(* IEC 61131-3 sources: daoli-st-library/DL_Base (part 6) *)

(* ---- FC_DL_MapRangeIntQuant.st ---- *)
(*
  FC_DL_MapRangeIntQuant —— 量程映射加整数量化，步长加四舍五入
  分类：DL_Base | 复杂度：2 | 轮次：R86
  开源溯源：道莅原创（clean-room 自研，纯 IEC 61131-3 通用算法），无外部代码引用
  许可证：MIT
  职责：先把输入线性映射到输出量程（输入越界钳位），再按 fStep 步长量化到整数刻度：
        nTick = round(mapped / step)，fOut = nTick * step；fTick 为量化后的整数刻度。
  契约：fIn 输入、fInMin/fInMax 输入端点、fOutMin/fOutMax 输出端点、fStep 步长（必须 > 0）；
        fOut 量化结果 [输出量程单位]、fTick 整数刻度；返回 TRUE 表示可信。
  边界：① 步长零 / 负值前置判（除零防护）；② 量程退化校验（容差 DL_MQ_EPS）；
        ③ 六个浮点入参逐一非有限闸；④ 转整前对刻度做 ±1.0E6 上限兜底，避免 LREAL_TO_DINT 越域；
        ⑤ 零全局、零物理地址、零库件依赖。
*)
FUNCTION FC_DL_MapRangeIntQuant : BOOL
VAR_INPUT
    fIn     : LREAL := 0.0;            // 输入值 [输入量程单位] / The input value
    fInMin  : LREAL := 0.0;            // 输入量程下端点 [输入量程单位] / The input range low end
    fInMax  : LREAL := 100.0;          // 输入量程上端点 [输入量程单位] / The input range high end
    fOutMin : LREAL := 0.0;            // 输出量程下端点 [输出量程单位] / The output range low end
    fOutMax : LREAL := 100.0;          // 输出量程上端点 [输出量程单位] / The output range high end
    fStep   : LREAL := 1.0;            // 量化步长（必须 > 0） [输出量程单位] / The quantisation step
END_VAR
VAR_OUTPUT
    fOut  : LREAL;                     // 量化后的结果 [输出量程单位] / The quantised result
    fTick : LREAL;                     // 量化后的整数刻度值 [刻度] / The integer tick value as a real
END_VAR
VAR
    xBad     : BOOL;                   // 参数非法标志 [—] / The parameter invalid flag
    fInSpan  : LREAL;                  // 输入量程跨度 [输入量程单位] / The input span
    fMapped  : LREAL;                  // 未量化的映射值 [输出量程单位] / The mapped value
    fTicks   : LREAL;                  // 未取整的刻度 [刻度] / The raw tick count
    diTick   : DINT;                   // 四舍五入后的整数刻度 [刻度] / The rounded tick count
END_VAR
VAR CONSTANT
    DL_MQ_EPS  : LREAL := 1.0E-9;      // 浮点比较容差 [-] / The floating point comparison tolerance
    DL_MQ_INF  : LREAL := 1.0E30;      // 非有限 / 越界判据上限 [-] / The magnitude gate
    DL_MQ_TICK : LREAL := 1.0E6;       // 转整前的刻度上限兜底 [刻度] / The tick guard before conversion
    DL_MQ_HALF : LREAL := 0.5;         // 四舍五入偏置 [-] / The rounding bias
    DL_MQ_Z    : LREAL := 0.0;         // 浮点零常量 [-] / The floating point zero constant
END_VAR

FC_DL_MapRangeIntQuant := FALSE;                          // 返回值预置假 / preset the return false
fOut := fOutMin;                                          // 输出预置为输出下端点哨兵 / preset the low end sentinel
fTick := DL_MQ_Z;                                         // 刻度预置零 [刻度] / preset the tick zero
xBad := FALSE;                                            // 非法标志预置假 / preset the invalid flag false
IF (fIn <> fIn) OR (ABS(fIn) > DL_MQ_INF) THEN            // 输入非有限闸 / the input gate
    xBad := TRUE;                                         // 置非法标志 / raise the invalid flag
END_IF
IF (fInMin <> fInMin) OR (ABS(fInMin) > DL_MQ_INF) THEN   // 输入下端非有限闸 / the input low end gate
    xBad := TRUE;                                         // 置非法标志 / raise the invalid flag
END_IF
IF (fInMax <> fInMax) OR (ABS(fInMax) > DL_MQ_INF) THEN   // 输入上端非有限闸 / the input high end gate
    xBad := TRUE;                                         // 置非法标志 / raise the invalid flag
END_IF
IF (fOutMin <> fOutMin) OR (ABS(fOutMin) > DL_MQ_INF) THEN // 输出下端非有限闸 / the output low end gate
    xBad := TRUE;                                         // 置非法标志 / raise the invalid flag
END_IF
IF (fOutMax <> fOutMax) OR (ABS(fOutMax) > DL_MQ_INF) THEN // 输出上端非有限闸 / the output high end gate
    xBad := TRUE;                                         // 置非法标志 / raise the invalid flag
END_IF
IF (fStep <> fStep) OR (ABS(fStep) > DL_MQ_INF) THEN      // 步长非有限闸 / the step gate
    xBad := TRUE;                                         // 置非法标志 / raise the invalid flag
END_IF
IF fStep <= DL_MQ_EPS THEN                                // 步长非正（除零防护） / the step is not positive
    xBad := TRUE;                                         // 置非法标志 / raise the invalid flag
END_IF
fInSpan := fInMax - fInMin;                               // 输入量程跨度 [输入量程单位] / the input span
IF ABS(fInSpan) < DL_MQ_EPS THEN                          // 输入量程退化（除零防护） / the degenerate input span
    xBad := TRUE;                                         // 置非法标志 / raise the invalid flag
END_IF
IF NOT xBad THEN                                          // 参数全通过才映射量化 / map and quantise when all pass
    fMapped := fIn;                                       // 输入接管 [输入量程单位] / take the input value
    IF fInSpan > DL_MQ_Z THEN                             // 正常量程方向 / the normal direction
        IF fMapped < fInMin THEN                          // 低于下端点 / below the low end
            fMapped := fInMin;                            // 钳到下端点 [输入量程单位] / clamp to the low end
        END_IF
        IF fMapped > fInMax THEN                          // 高于上端点 / above the high end
            fMapped := fInMax;                            // 钳到上端点 [输入量程单位] / clamp to the high end
        END_IF
    ELSE                                                  // 反向量程 / the reversed direction
        IF fMapped > fInMin THEN                          // 高于下端点 / above the low end
            fMapped := fInMin;                            // 钳到下端点 [输入量程单位] / clamp to the low end
        END_IF
        IF fMapped < fInMax THEN                          // 低于上端点 / below the high end
            fMapped := fInMax;                            // 钳到上端点 [输入量程单位] / clamp to the high end
        END_IF
    END_IF
    fMapped := fOutMin + ((fMapped - fInMin) / fInSpan) * (fOutMax - fOutMin); // 线性映射（分母已证非零）
    fTicks := fMapped / fStep;                            // 换算成刻度数（步长已证正） [刻度] / the raw tick count
    IF fTicks > DL_MQ_TICK THEN                           // 刻度上越界，转整前兜底 / the positive tick guard
        fTicks := DL_MQ_TICK;                             // 钳到刻度上限 [刻度] / clamp the tick count
    END_IF
    IF fTicks < -DL_MQ_TICK THEN                          // 刻度下越界，转整前兜底 / the negative tick guard
        fTicks := -DL_MQ_TICK;                            // 钳到刻度下限 [刻度] / clamp the tick count
    END_IF
    IF fTicks >= DL_MQ_HALF THEN                          // 非负四舍五入 / non negative rounding
        diTick := LREAL_TO_DINT(fTicks + DL_MQ_HALF);     // 加半后截断 [刻度] / add a half then truncate
    ELSIF fTicks <= -DL_MQ_HALF THEN                      // 非正四舍五入 / non positive rounding
        diTick := LREAL_TO_DINT(fTicks - DL_MQ_HALF);     // 减半后截断 [刻度] / subtract a half then truncate
    ELSE
        diTick := 0;                                      // 近零带归零 [刻度] / the near zero band
    END_IF
    fTick := DINT_TO_LREAL(diTick);                       // 整数刻度出口 [刻度] / publish the integer tick
    fOut := fTick * fStep;                                // 量化结果还原 [输出量程单位] / restore the quantised value
    FC_DL_MapRangeIntQuant := TRUE;                       // 量化成功 / the quantisation succeeded
ELSE
    fOut := fOutMin;                                      // 非法参数输出下端点哨兵 [输出量程单位] / the sentinel
    fTick := DL_MQ_Z;                                     // 刻度输出零哨兵 [刻度] / the tick sentinel
    FC_DL_MapRangeIntQuant := FALSE;                      // 结果不可信 / the result is not valid
END_IF
END_FUNCTION

(* ---- FC_DL_MapRangeInverseSolve.st ---- *)
(*
  FC_DL_MapRangeInverseSolve —— 由工程值反解原始量程值，含钳位
  分类：DL_Base | 复杂度：2 | 轮次：R86
  开源溯源：道莅原创（clean-room 自研，纯 IEC 61131-3 通用算法），无外部代码引用
  许可证：MIT
  职责：正向映射 out = fOutMin + (in - fInMin)/(fInMax - fInMin) * (fOutMax - fOutMin) 的逆解：
        raw = fInMin + (fOut - fOutMin) * (fInMax - fInMin) / (fOutMax - fOutMin)。
  契约：fEng 工程值输入 [输出量程单位]、fInMin/fInMax 原始量程端点、fOutMin/fOutMax 工程量程端点；
        fRaw 反解结果 [原始量程单位]（钳在原始量程内）；返回 TRUE 表示可信。
  边界：① 除零防护：分母 fOutSpan 过退化闸后才做除法；② 反解结果按原始量程钳位；
        ③ 五个浮点入参逐一非有限闸；④ 零全局、零物理地址、零库件依赖。
*)
FUNCTION FC_DL_MapRangeInverseSolve : BOOL
VAR_INPUT
    fEng    : LREAL := 0.0;            // 工程值输入 [输出量程单位] / The engineering value input
    fInMin  : LREAL := 0.0;            // 原始量程下端点 [原始量程单位] / The raw range low end
    fInMax  : LREAL := 100.0;          // 原始量程上端点 [原始量程单位] / The raw range high end
    fOutMin : LREAL := 0.0;            // 工程量程下端点 [输出量程单位] / The engineering range low end
    fOutMax : LREAL := 100.0;          // 工程量程上端点 [输出量程单位] / The engineering range high end
END_VAR
VAR_OUTPUT
    fRaw : LREAL;                      // 反解结果 [原始量程单位] / The solved raw value
END_VAR
VAR
    xBad      : BOOL;                  // 参数非法标志 [—] / The parameter invalid flag
    fEngClamp : LREAL;                 // 钳位后的工程值 [输出量程单位] / The clamped engineering value
    fOutSpan  : LREAL;                 // 工程量程跨度 [输出量程单位] / The engineering span
    fInSpan   : LREAL;                 // 原始量程跨度 [原始量程单位] / The raw span
    fRawCalc  : LREAL;                 // 未钳位的反解结果 [原始量程单位] / The unclamped solved value
END_VAR
VAR CONSTANT
    DL_MI_EPS : LREAL := 1.0E-9;       // 浮点比较容差 [-] / The floating point comparison tolerance
    DL_MI_INF : LREAL := 1.0E30;       // 非有限 / 越界判据上限 [-] / The magnitude gate
    DL_MI_Z   : LREAL := 0.0;          // 浮点零常量 [-] / The floating point zero constant
END_VAR

FC_DL_MapRangeInverseSolve := FALSE;                      // 返回值预置假 / preset the return false
fRaw := fInMin;                                           // 输出预置为原始量程下端点哨兵 / preset the raw low end sentinel
xBad := FALSE;                                            // 非法标志预置假 / preset the invalid flag false
IF (fEng <> fEng) OR (ABS(fEng) > DL_MI_INF) THEN         // 工程值非有限闸 / the engineering value gate
    xBad := TRUE;                                         // 置非法标志 / raise the invalid flag
END_IF
IF (fInMin <> fInMin) OR (ABS(fInMin) > DL_MI_INF) THEN   // 原始下端非有限闸 / the raw low end gate
    xBad := TRUE;                                         // 置非法标志 / raise the invalid flag
END_IF
IF (fInMax <> fInMax) OR (ABS(fInMax) > DL_MI_INF) THEN   // 原始上端非有限闸 / the raw high end gate
    xBad := TRUE;                                         // 置非法标志 / raise the invalid flag
END_IF
IF (fOutMin <> fOutMin) OR (ABS(fOutMin) > DL_MI_INF) THEN // 工程下端非有限闸 / the engineering low end gate
    xBad := TRUE;                                         // 置非法标志 / raise the invalid flag
END_IF
IF (fOutMax <> fOutMax) OR (ABS(fOutMax) > DL_MI_INF) THEN // 工程上端非有限闸 / the engineering high end gate
    xBad := TRUE;                                         // 置非法标志 / raise the invalid flag
END_IF
fOutSpan := fOutMax - fOutMin;                            // 工程量程跨度 [输出量程单位] / the engineering span
fInSpan := fInMax - fInMin;                               // 原始量程跨度 [原始量程单位] / the raw span
IF ABS(fOutSpan) < DL_MI_EPS THEN                         // 工程跨度退化（除零防护） / the degenerate engineering span
    xBad := TRUE;                                         // 置非法标志 / raise the invalid flag
END_IF
IF NOT xBad THEN                                          // 参数全通过才反解 / solve only when all parameters pass
    fEngClamp := fEng;                                    // 工程值接管 [输出量程单位] / take the engineering value
    IF fOutSpan > DL_MI_Z THEN                            // 正常方向 / the normal direction
        IF fEngClamp < fOutMin THEN                       // 低于工程下端点 / below the engineering low end
            fEngClamp := fOutMin;                         // 钳到工程下端点 [输出量程单位] / clamp to the low end
        END_IF
        IF fEngClamp > fOutMax THEN                       // 高于工程上端点 / above the engineering high end
            fEngClamp := fOutMax;                         // 钳到工程上端点 [输出量程单位] / clamp to the high end
        END_IF
    ELSE                                                  // 反向工程跨度 / the reversed engineering span
        IF fEngClamp > fOutMin THEN                       // 高于工程下端点 / above the engineering low end
            fEngClamp := fOutMin;                         // 钳到工程下端点 [输出量程单位] / clamp to the low end
        END_IF
        IF fEngClamp < fOutMax THEN                       // 低于工程上端点 / below the engineering high end
            fEngClamp := fOutMax;                         // 钳到工程上端点 [输出量程单位] / clamp to the high end
        END_IF
    END_IF
    fRawCalc := fInMin + ((fEngClamp - fOutMin) / fOutSpan) * fInSpan; // 反解（分母已证非零） [原始量程单位]
    IF fInMax >= fInMin THEN                              // 原始量程正常方向 / the normal raw direction
        IF fRawCalc < fInMin THEN                         // 反解低于原始下端点 / below the raw low end
            fRawCalc := fInMin;                           // 钳到原始下端点 [原始量程单位] / clamp to the low end
        END_IF
        IF fRawCalc > fInMax THEN                         // 反解高于原始上端点 / above the raw high end
            fRawCalc := fInMax;                           // 钳到原始上端点 [原始量程单位] / clamp to the high end
        END_IF
    ELSE                                                  // 原始量程反向 / the reversed raw range
        IF fRawCalc > fInMin THEN                         // 反解高于原始下端点 / above the raw low end
            fRawCalc := fInMin;                           // 钳到原始下端点 [原始量程单位] / clamp to the low end
        END_IF
        IF fRawCalc < fInMax THEN                         // 反解低于原始上端点 / below the raw high end
            fRawCalc := fInMax;                           // 钳到原始上端点 [原始量程单位] / clamp to the high end
        END_IF
    END_IF
    fRaw := fRawCalc;                                     // 反解结果出口 [原始量程单位] / publish the solved value
    FC_DL_MapRangeInverseSolve := TRUE;                   // 反解成功 / the solve succeeded
ELSE
    fRaw := fInMin;                                       // 非法参数输出原始下端点哨兵 [原始量程单位] / the sentinel
    FC_DL_MapRangeInverseSolve := FALSE;                  // 结果不可信 / the result is not valid
END_IF
END_FUNCTION

(* ---- FC_DL_MapRangePiecewise3.st ---- *)
(*
  FC_DL_MapRangePiecewise3 —— 三段折线映射，分段斜率加断点连续校验
  分类：DL_Base | 复杂度：2 | 轮次：R86
  开源溯源：道莅原创（clean-room 自研，纯 IEC 61131-3 通用算法），无外部代码引用
  许可证：MIT
  职责：由 4 个断点（afX 单调递增）与对应 4 个输出值构造三段折线，按输入落在哪一段做线性插值；
        断点单调性即保证折线在断点处连续（左段右端值 = 右段左端值 = afY[i]）。
  契约：fIn 输入、afX 断点横坐标（必须严格递增）、afY 断点纵坐标；fOut 折线输出；返回 TRUE 表示可信。
  边界：① 断点严格递增校验（容差 DL_MW_EPS），否则判非法；② 所有断点与输入做非有限闸；
        ③ 输入越两端断点时钳到端点（不外插）；④ 除零防护：段跨度经单调性闸后恒 > 0；
        ⑤ 零全局、零物理地址、零库件依赖；数组为显式定长（R15）。
*)
FUNCTION FC_DL_MapRangePiecewise3 : BOOL
VAR_INPUT
    fIn  : LREAL := 0.0;                             // 输入值 [输入量程单位] / The input value
    afX  : ARRAY[0..3] OF LREAL;                     // 四个断点横坐标（严格递增） [输入量程单位] / The breakpoints
    afY  : ARRAY[0..3] OF LREAL;                     // 四个断点纵坐标 [输出量程单位] / The breakpoint outputs
END_VAR
VAR_OUTPUT
    fOut  : LREAL;                                   // 折线输出 [输出量程单位] / The piecewise output
    nSeg  : INT;                                     // 命中段号（0..2） [下标] / The hit segment index
END_VAR
VAR
    xBad  : BOOL;                                    // 参数非法标志 [—] / The parameter invalid flag
    xFound : BOOL;                                   // 命中段查找标志 [—] / The hit segment search flag
    i     : INT;                                     // 遍历索引 [下标] / The traversal index
    k     : INT;                                     // 命中段索引 [下标] / The hit segment index
    fSpan : LREAL;                                   // 命中段的横坐标跨度 [输入量程单位] / The segment span
END_VAR
VAR CONSTANT
    DL_MW_EPS  : LREAL := 1.0E-9;                    // 浮点比较容差 [-] / The floating point comparison tolerance
    DL_MW_INF  : LREAL := 1.0E30;                    // 非有限 / 越界判据上限 [-] / The magnitude gate
    DL_MW_Z    : LREAL := 0.0;                       // 浮点零常量 [-] / The floating point zero constant
    DL_MW_N    : INT := 3;                           // 折线段数 [段] / The number of segments
    DL_MW_I0   : INT := 0;                           // 下标零 [下标] / The index zero
END_VAR

FC_DL_MapRangePiecewise3 := FALSE;                    // 返回值预置假 / preset the return false
fOut := DL_MW_Z;                                      // 输出预置零哨兵 / preset the zero sentinel
nSeg := DL_MW_I0;                                     // 段号预置零 [下标] / preset the segment index zero
xBad := FALSE;                                        // 非法标志预置假 / preset the invalid flag false
IF (fIn <> fIn) OR (ABS(fIn) > DL_MW_INF) THEN        // 输入非有限闸 / the input gate
    xBad := TRUE;                                     // 置非法标志 / raise the invalid flag
END_IF
FOR i := DL_MW_I0 TO DL_MW_N DO                       // 四个断点逐一校验 / check every breakpoint
    IF (afX[i] <> afX[i]) OR (ABS(afX[i]) > DL_MW_INF) THEN // 横坐标非有限 / the abscissa is not finite
        xBad := TRUE;                                 // 置非法标志 / raise the invalid flag
    END_IF
    IF (afY[i] <> afY[i]) OR (ABS(afY[i]) > DL_MW_INF) THEN // 纵坐标非有限 / the ordinate is not finite
        xBad := TRUE;                                 // 置非法标志 / raise the invalid flag
    END_IF
END_FOR
FOR i := DL_MW_I0 TO DL_MW_N - 1 DO                   // 相邻断点严格递增校验 / strictly increasing check
    IF (afX[i + 1] - afX[i]) < DL_MW_EPS THEN         // 跨度非正（含重合断点） / a non positive span
        xBad := TRUE;                                 // 置非法标志 / raise the invalid flag
    END_IF
END_FOR
IF NOT xBad THEN                                      // 参数全通过才插值 / interpolate when all parameters pass
    IF fIn <= afX[DL_MW_I0] THEN                      // 低于最低断点，钳到端点 / below the lowest breakpoint
        fOut := afY[DL_MW_I0];                        // 取最低断点输出 [输出量程单位] / take the lowest output
        nSeg := DL_MW_I0;                             // 段号记零 [下标] / the segment index is zero
    ELSIF fIn >= afX[DL_MW_N] THEN                    // 高于最高断点，钳到端点 / above the highest breakpoint
        fOut := afY[DL_MW_N];                         // 取最高断点输出 [输出量程单位] / take the highest output
        nSeg := DL_MW_N - 1;                          // 段号记末段 [下标] / the last segment index
    ELSE
        k := DL_MW_I0;                                // 段索引从零起 / the segment index starts at zero
        xFound := FALSE;                              // 命中标志预置假 / preset the hit flag false
        WHILE (k <= DL_MW_N - 1) AND NOT xFound DO    // 显式递增查找命中段（有界） / find the hit segment
            IF fIn < afX[k + 1] THEN                  // 落在第 k 段内 / inside the k th segment
                xFound := TRUE;                       // 置命中标志 / raise the hit flag
            ELSE
                k := k + 1;                           // 继续下一段 / advance to the next segment
            END_IF
        END_WHILE
        IF k > DL_MW_N - 1 THEN                       // 命中段上越界兜底 / the hit index fallback
            k := DL_MW_N - 1;                         // 钳到末段 [下标] / clamp to the last segment
        END_IF
        fSpan := afX[k + 1] - afX[k];                 // 命中段跨度（已证 > 容差） [输入量程单位] / the segment span
        fOut := afY[k] + ((fIn - afX[k]) / fSpan) * (afY[k + 1] - afY[k]); // 段内线性插值 [输出量程单位]
        nSeg := k;                                    // 段号出口 [下标] / publish the hit segment
    END_IF
    FC_DL_MapRangePiecewise3 := TRUE;                 // 插值成功 / the interpolation succeeded
ELSE
    fOut := DL_MW_Z;                                  // 非法参数输出零哨兵 [输出量程单位] / the sentinel
    FC_DL_MapRangePiecewise3 := FALSE;                // 结果不可信 / the result is not valid
END_IF
END_FUNCTION

(* ---- FC_DL_MapRangeSatOut.st ---- *)
(*
  FC_DL_MapRangeSatOut —— 输入量程映射后对输出独立饱和限幅
  分类：DL_Base | 复杂度：2 | 轮次：R86
  开源溯源：道莅原创（clean-room 自研，纯 IEC 61131-3 通用算法），无外部代码引用
  许可证：MIT
  职责：先做 [fInMin, fInMax] → [fOutMin, fOutMax] 的线性映射（输入先钳到量程），
        再把映射结果独立钳到执行机构允许的 [fSatMin, fSatMax]（该区间可比输出量程更窄）。
  契约：fIn 输入、fInMin/fInMax 输入端点、fOutMin/fOutMax 输出端点、fSatMin/fSatMax 输出饱和限；
        fOut 结果；xSat 报告输出侧发生饱和；返回 TRUE 表示可信。
  边界：① 输入量程与饱和区间双退化校验（容差 DL_MS_EPS）；② 八个浮点入参逐一非有限闸；
        ③ 除零防护：除以 fInSpan 前已过退化闸；④ 零全局、零物理地址、零库件依赖。
*)
FUNCTION FC_DL_MapRangeSatOut : BOOL
VAR_INPUT
    fIn     : LREAL := 0.0;            // 输入值 [输入量程单位] / The input value
    fInMin  : LREAL := 0.0;            // 输入量程下端点 [输入量程单位] / The input range low end
    fInMax  : LREAL := 100.0;          // 输入量程上端点 [输入量程单位] / The input range high end
    fOutMin : LREAL := 0.0;            // 输出量程下端点 [输出量程单位] / The output range low end
    fOutMax : LREAL := 100.0;          // 输出量程上端点 [输出量程单位] / The output range high end
    fSatMin : LREAL := 0.0;            // 输出饱和下限 [输出量程单位] / The output saturation low limit
    fSatMax : LREAL := 100.0;          // 输出饱和上限 [输出量程单位] / The output saturation high limit
END_VAR
VAR_OUTPUT
    fOut : LREAL;                      // 结果（含输出侧饱和） [输出量程单位] / The saturated result
    xSat : BOOL;                       // 输出侧发生饱和 [—] / The output stage saturated
END_VAR
VAR
    xBad      : BOOL;                  // 参数非法标志 [—] / The parameter invalid flag
    fInClamp  : LREAL;                 // 钳位后的输入 [输入量程单位] / The clamped input
    fInSpan   : LREAL;                 // 输入量程跨度 [输入量程单位] / The input span
    fMapped   : LREAL;                 // 未限幅的映射结果 [输出量程单位] / The mapped value before limiting
END_VAR
VAR CONSTANT
    DL_MS_EPS : LREAL := 1.0E-9;       // 浮点比较容差 [-] / The floating point comparison tolerance
    DL_MS_INF : LREAL := 1.0E30;       // 非有限 / 越界判据上限 [-] / The magnitude gate
    DL_MS_Z   : LREAL := 0.0;          // 浮点零常量 [-] / The floating point zero constant
END_VAR

FC_DL_MapRangeSatOut := FALSE;                            // 返回值预置假 / preset the return false
fOut := fOutMin;                                          // 输出预置为输出下端点哨兵 / preset the low end sentinel
xSat := FALSE;                                            // 饱和标志预置假 / preset the saturation flag false
xBad := FALSE;                                            // 非法标志预置假 / preset the invalid flag false
IF (fIn <> fIn) OR (ABS(fIn) > DL_MS_INF) THEN            // 输入非有限闸 / the input gate
    xBad := TRUE;                                         // 置非法标志 / raise the invalid flag
END_IF
IF (fInMin <> fInMin) OR (ABS(fInMin) > DL_MS_INF) THEN   // 输入下端非有限闸 / the input low end gate
    xBad := TRUE;                                         // 置非法标志 / raise the invalid flag
END_IF
IF (fInMax <> fInMax) OR (ABS(fInMax) > DL_MS_INF) THEN   // 输入上端非有限闸 / the input high end gate
    xBad := TRUE;                                         // 置非法标志 / raise the invalid flag
END_IF
IF (fOutMin <> fOutMin) OR (ABS(fOutMin) > DL_MS_INF) THEN // 输出下端非有限闸 / the output low end gate
    xBad := TRUE;                                         // 置非法标志 / raise the invalid flag
END_IF
IF (fOutMax <> fOutMax) OR (ABS(fOutMax) > DL_MS_INF) THEN // 输出上端非有限闸 / the output high end gate
    xBad := TRUE;                                         // 置非法标志 / raise the invalid flag
END_IF
IF (fSatMin <> fSatMin) OR (ABS(fSatMin) > DL_MS_INF) THEN // 饱和下限非有限闸 / the saturation low gate
    xBad := TRUE;                                         // 置非法标志 / raise the invalid flag
END_IF
IF (fSatMax <> fSatMax) OR (ABS(fSatMax) > DL_MS_INF) THEN // 饱和上限非有限闸 / the saturation high gate
    xBad := TRUE;                                         // 置非法标志 / raise the invalid flag
END_IF
fInSpan := fInMax - fInMin;                               // 输入量程跨度 [输入量程单位] / the input span
IF ABS(fInSpan) < DL_MS_EPS THEN                          // 输入量程退化（除零防护） / the degenerate input span
    xBad := TRUE;                                         // 置非法标志 / raise the invalid flag
END_IF
IF fSatMax < fSatMin THEN                                 // 饱和区间倒置 / the saturated band is inverted
    xBad := TRUE;                                         // 置非法标志 / raise the invalid flag
END_IF
IF NOT xBad THEN                                          // 参数全通过才映射 / map only when all parameters pass
    fInClamp := fIn;                                      // 输入接管 [输入量程单位] / take the input value
    IF fInSpan > DL_MS_Z THEN                             // 正常量程方向 / the normal direction
        IF fInClamp < fInMin THEN                         // 低于下端点 / below the low end
            fInClamp := fInMin;                           // 钳到下端点 [输入量程单位] / clamp to the low end
        END_IF
        IF fInClamp > fInMax THEN                         // 高于上端点 / above the high end
            fInClamp := fInMax;                           // 钳到上端点 [输入量程单位] / clamp to the high end
        END_IF
    ELSE                                                  // 反向量程 / the reversed direction
        IF fInClamp > fInMin THEN                         // 高于下端点 / above the low end
            fInClamp := fInMin;                           // 钳到下端点 [输入量程单位] / clamp to the low end
        END_IF
        IF fInClamp < fInMax THEN                         // 低于上端点 / below the high end
            fInClamp := fInMax;                           // 钳到上端点 [输入量程单位] / clamp to the high end
        END_IF
    END_IF
    fMapped := fOutMin + ((fInClamp - fInMin) / fInSpan) * (fOutMax - fOutMin); // 线性映射（分母已证非零）
    fOut := fMapped;                                      // 映射值接入输出侧限幅 [输出量程单位] / take the mapped value
    IF fMapped > fSatMax THEN                             // 输出侧上饱和 / the output stage saturates high
        fOut := fSatMax;                                  // 钳到饱和上限 [输出量程单位] / clamp to the high limit
        xSat := TRUE;                                     // 置饱和标志 [—] / raise the saturation flag
    END_IF
    IF fMapped < fSatMin THEN                             // 输出侧下饱和 / the output stage saturates low
        fOut := fSatMin;                                  // 钳到饱和下限 [输出量程单位] / clamp to the low limit
        xSat := TRUE;                                     // 置饱和标志 [—] / raise the saturation flag
    END_IF
    FC_DL_MapRangeSatOut := TRUE;                         // 映射成功 / the mapping succeeded
ELSE
    fOut := fOutMin;                                      // 非法参数输出下端点哨兵 [输出量程单位] / the sentinel
    FC_DL_MapRangeSatOut := FALSE;                        // 结果不可信 / the result is not valid
END_IF
END_FUNCTION

(* ---- FC_DL_MaskCompare.st ---- *)
(*==============================================================================
 * 组件名称 (Component)  : FC_DL_MaskCompare
 * 所属子库 (Sublibrary) : DL_Base
 * 归属目录 (Directory)  : C:\Library\DL_Base
 * 当前版本 (Version)    : 1.0.0
 * 分类/来源标签         : 函数（FUNCTION）· 纯函数 · 状态字掩码比较与差异定位
 *                         lgf-comparator / lgf-bitlogic / mask-compare
 * 兼容性   (Platform)   : CODESYS 3.5 / TwinCAT 3 / 汇川 InoProShop / 施耐德
 *                         Machine Expert；仅用 Standard.library 的 SHL / SHR /
 *                         AND / XOR，无厂商位访问方言，无实例依赖
 * 功能一句话 (Summary)  : 判「值按掩码比较是否等于期望」，并给出差异位图、差异
 *                         位数与首个差异位号，供报警直接定位到具体那一位。
 * 功能描述 (Function)   : 核心判据为「值与期望各自按掩码相与后判等」。掩码为 0 的位
 *                         不参与比较（don't-care 位），位宽参数把高于 nWidth 减 1 的
 *                         位排除在比较之外（只比低 n 位）。典型现场用途：变频器状态
 *                         字只看「运行、故障、就绪」三位的组合、远程 IO 模块状态字
 *                         忽略保留位后的整字比对、多轴使能位图的期望态一致性检查、
 *                         以及报警诊断时直接报出「差在第几位」而不是只说「不匹配」。
 * 与既有件边界 (Boundary): FC_DL_BitFieldExtract 是「取一段」（把位段取出后由调用方
 *                         自行比较）；FB_DL_StatusWordSegDecoder 是「段表批量解码」
 *                         （把状态字按段拆成多个语义位）；本件是「判等 + 差异定位」，
 *                         一次调用既回答「是否匹配」又回答「差在哪几位」。三者互补，
 *                         不互相替代。
 * 设计要点 (Key notes)  : ① 掩码与位宽两重屏蔽严格串联：先按位宽裁出有效位域，再与
 *                           调用方掩码相与，两道屏蔽同时生效，不存在「宽掩码压过窄位宽」
 *                           的漏判；
 *                         ② 位宽 32 走全一常量分支，禁止 SHL 移位量等于位宽（部分
 *                           编译器对此属未定义行为）；
 *                         ③ 差异位号由低位向高位扫描，报「最低的那个差异位」，与现场
 *                           按位号读状态字的习惯一致；
 *                         ④ 纯函数：无内部状态、无跨周期残留，同入参同结果。
 *
 * 【验收向量 / Acceptance vectors】
 *   V1  值 16#1234_5678、期望 16#0034_5678、掩码 16#00FF_FFFF
 *       → 返回真、差异位图 0、差异位数 0、首差位 负 1（高 8 位被掩掉，不参与）
 *   V2  同 V1 但期望改 16#0034_5670 → 返回假、差异位图 16#0000_0008、
 *       差异位数 1、首差位 3
 *   V3  V-A 域外：位宽 0 → 返回假、码 0220、差异位图 0（不输出脏位图）
 *   V4  V-B 边界：位宽 32、掩码全一、值 0、期望 16#8000_0000
 *       → 返回假、首差位 31（验证 32 位常量掩码路径，不做按位宽移位）
 *   V5  位宽 5、掩码 16#FFFF_FFFF、值 16#0000_0020、期望 0
 *       → 返回真、差异位图 0（第 5 位及以上被位宽裁掉，越界位不参与比较）
 *   V6  掩码 0 → 返回真、码 0140（恒匹配，提示掩码没生效）
 *
 * 开源溯源 (Origin)     : 来源标签 lgf-comparator 与 lgf-bitlogic。LGF（Libre
 *                         Graphical Framework）为免费闭源发布的公开函数库手册，
 *                         本件仅借鉴其「二进制掩码比较」块的语义域（值、期望、掩码
 *                         三引脚）与比较器组「单值、区间、掩码」的分类粒度；许可证
 *                         按其发布方条款仅作分类参考，本件零代码行、零注释、零数据
 *                         结构引用，属 clean-room 独立实现，不构成衍生作品。
 * 码位说明 (Codes)      : 信息 16#0001_013F 位宽已钳到 32 ｜ 16#0001_0140 掩码为 0
 *                         故障 16#0001_0220 位宽非法。取号见本轮规格 §3.2，与位段族
 *                         0125 到 013E 区间不重叠。
 * 依赖说明 (Depends)    : 无 DL_ 内部依赖；仅 Standard.library 的 SHL / SHR / AND /
 *                         XOR 与 INT_TO_UDINT 显式转换。
 * 镜像量清单 (R38)      : 本件无锁存副本，差异位图与差异位数都由同一份本拍差值导出，
 *                         不存在锁存量与实时量混用面。
 * 红线自检 (Redline)    : 零全局变量表依赖 ｜ 零外部变量声明 ｜ 零物理地址直写
 *                         纯 IEC 61131-3 ｜ 无除法故无除零面 ｜ 位宽 32 走常量分支
 *                         全变量双语同行注释 ｜ 状态机 N/A（纯函数）｜ 无定时器实例
 * 修订历史 (Revision)   : 2026-11-15  v1.0.0  首版入库（Round 13 · 泳道 B 位段族收口）
 *============================================================================*)

(*==============================================================================
 * 双重屏蔽示意 (Double masking)：
 *   位宽 5、掩码全一、值 16#0000_0020、期望 0
 *   第一步按位宽裁出低位域 16#0000_001F
 *   第二步与掩码相与仍为 16#0000_001F
 *   值域为 0、期望域为 0，差为 0，返回真；第 5 位虽然置位但不在契约位宽内
 *   若掩码改为 16#0000_0020 而位宽仍是 5，有效掩码变成 0，属「掩码被位宽吃掉」，
 *   此时按恒匹配处理并给出 0140，提示调用方掩码与位宽矛盾
 *============================================================================*)

FUNCTION FC_DL_MaskCompare : BOOL
VAR_INPUT
    uValue  : DWORD;                    // 待比较值 [位串] / Value under test
    uExpect : DWORD;                    // 期望值 [位串] / Expected value
    uMask   : DWORD := 16#FFFF_FFFF;    // 参与比较的位，1 参与比较、0 不关心 [位串] / Care mask, one means compare
    nWidth  : INT := 32;                // 有效位宽 [bit]，域 1 到 32 / Effective width, 1 to 32
END_VAR
VAR_OUTPUT
    uDiffBits  : DWORD;                 // 差异位图，已按位宽与掩码双重屏蔽 [位串] / Difference bitmap after both masks
    nDiffCount : INT;                   // 差异位数 [个]，域 0 到 32 / Difference bit count, 0 to 32
    nFirstDiff : INT;                   // 首个差异位号 [bit]，域 0 到 31，无差异为负 1 / First differing bit, minus one when none
    uErrorId   : UDINT;                 // 事件码，0 表示无事件 / Event code, zero means none
END_VAR
VAR
    nW         : INT;                   // 钳位后的有效位宽 [bit] / Clamped effective width
    uWidthMask : DWORD;                 // 位宽掩码，低 nW 位为 1 [位串] / Width mask with the low nW bits set
    uMaskEff   : DWORD;                 // 生效掩码，位宽掩码与调用方掩码相与 [位串] / Effective mask combining width and caller mask
    uDiff      : DWORD;                 // 值与期望按生效掩码异或的结果 [位串] / XOR result under the effective mask
    uScan      : DWORD;                 // 扫描副本，逐位右移 [位串] / Shifting scan copy
    nI         : INT;                   // 位扫描下标 [bit]，固定 0 到 31 / Bit scan index, fixed 0 to 31
    nCount     : INT;                   // 差异位计数累加 [个] / Running difference count
    nFirst     : INT;                   // 首个差异位累加，未命中保持负 1 / Running first differing bit, minus one when none
    uCode      : UDINT;                 // 码位暂存，出口单点写入 [码] / Code staging, written once at the exit
END_VAR
VAR CONSTANT
    DL_MC_MAXW    : INT := 32;                  // 最大位宽 [bit]，与位宽默认值一致 / Maximum width, matches the default width
    DL_MC_MASK32  : DWORD := 16#FFFF_FFFF;      // 满宽掩码常量，位宽 32 分支专用 [位串] / All ones mask for the 32 bit branch
    DL_MC_NONE    : INT := -1;                  // 无差异位号的表示值 [bit] / Sentinel for no differing bit
END_VAR

(*------------------------------------------------------------------------------
 * 段 1｜输出预置：差异类输出一律先归零，任何早退路径都不会留下脏位图
 *      Pre-set the difference outputs so early exits never publish stale bits
 *-----------------------------------------------------------------------------*)
FC_DL_MaskCompare := FALSE;
uDiffBits         := 16#0000_0000;
nDiffCount        := 0;
nFirstDiff        := DL_MC_NONE;
uErrorId          := 16#0000_0000;
uCode             := 16#0000_0000;
uDiff             := 16#0000_0000;
nCount            := 0;
nFirst            := DL_MC_NONE;

(*------------------------------------------------------------------------------
 * 段 2｜位宽闸门（边界 B1/B2）：小于 1 属逻辑错，早退；大于 32 钳位后照算
 *      Width gate: below one exits early, above thirty two is clamped
 *      位宽是契约参数，判错就把责任交回调用方，不用猜的值去凑结果
 *      The width is a contract parameter, guessing it would hide the configuration error
 *-----------------------------------------------------------------------------*)
IF nWidth < 1 THEN
    uErrorId := 16#0001_0220;   // 故障级：位宽非法，差异位图保持 0
    RETURN;
ELSIF nWidth > DL_MC_MAXW THEN
    nW    := DL_MC_MAXW;
    uCode := 16#0001_013F;      // 信息级：位宽已钳到 32
ELSE
    nW := nWidth;
END_IF

(*------------------------------------------------------------------------------
 * 段 3｜掩码构造（边界 B3）：位宽 32 用满一常量，其余用左移减一构造
 *      Mask construction: the full width case uses a constant, others shift minus one
 *      若在此处按位宽做移位，位宽 32 就会变成「移位量等于位宽」，属未定义行为
 *      Shifting by the full width here would be undefined behaviour on some compilers
 *-----------------------------------------------------------------------------*)
IF nW >= DL_MC_MAXW THEN
    uWidthMask := DL_MC_MASK32;
ELSE
    uWidthMask := SHL(DWORD#1, nW) - DWORD#1;
END_IF

uMaskEff := uMask AND uWidthMask;

(* 掩码为零属恒匹配：判据天然成立，但要提示调用方「掩码与位宽矛盾」
 * A zero mask matches anything, still worth telling the caller the mask is inert
 * 优先级低于位宽钳位码，故仅在未占用时写入
 * Lower priority than the clamp code above, written only when the slot is free *)
IF (uMaskEff = 16#0000_0000) AND (uCode = 16#0000_0000) THEN
    uCode := 16#0001_0140;
END_IF

(*------------------------------------------------------------------------------
 * 段 4｜判等与差异定位（边界 B4）：异或取差，逐位统计，先低后高
 *      Compare and locate: XOR the difference, then scan low bits first
 *      扫描固定 32 次、每次右移一位，移位量恒为 1，无动态移位风险
 *      The scan is a fixed thirty two passes shifting by one bit each time
 *-----------------------------------------------------------------------------*)
uDiff := (uValue XOR uExpect) AND uMaskEff;

IF uDiff = 16#0000_0000 THEN
    uDiffBits  := 16#0000_0000;
    nDiffCount := 0;
    nFirstDiff := DL_MC_NONE;
    FC_DL_MaskCompare := TRUE;          // 按契约位域完全一致 / Full match inside the contract bit field
ELSE
    uScan := uDiff;
    FOR nI := 0 TO (DL_MC_MAXW - 1) DO
        IF (uScan AND DWORD#1) = DWORD#1 THEN
            nCount := nCount + 1;
            IF nFirst = DL_MC_NONE THEN
                nFirst := nI;           // 首次命中即最低差异位 / The first hit is the lowest differing bit
            END_IF
        END_IF
        uScan := SHR(uScan, 1);
    END_FOR;
    uDiffBits  := uDiff;
    nDiffCount := nCount;
    nFirstDiff := nFirst;
    FC_DL_MaskCompare := FALSE;
END_IF

(*------------------------------------------------------------------------------
 * 段 5｜码位单点写入：全拍只写一次，优先级已在段 2 与段 3 排定
 *      Single write point for the code, the priority was settled above
 *-----------------------------------------------------------------------------*)
uErrorId := uCode;
END_FUNCTION

(* ---- FC_DL_PackBitsToWord.st ---- *)
(*==============================================================================
 * 组件名称 (Component)  : FC_DL_PackBitsToWord
 * 所属子库 (Sublibrary) : DL_Base
 * 当前版本 (Version)    : 1.0.0
 * 兼容性   (Platform)   : CODESYS 3.5 / TwinCAT 3 / 汇川 InoProShop / Machine Expert
 *                         仅用标准 SHL / OR / NOT，无任何厂商位写语法
 * 功能描述 (Function)   : 把 16 路离散 BOOL 状态打包成一个标准报警字 WORD，
 *                         供 Modbus / PROFINET 上传或写入设备状态字。
 *                         位序约定写死：数组索引 0 → bit0（LSB），不提供位序开关。
 *                         可选整体取反，适配低电平有效的报警点。
 * 开源溯源 (Origin)     : 原创实现。位序遵循 IEC 61131-3 位串类型"第 0 位为 LSB"规定。
 * 依赖     (Depends)    : 无 DL_ 内部依赖；无标准库功能块依赖
 *
 * 【uErrorId 显式豁免声明 / Explicit uErrorId exemption】
 *   本函数不设 uErrorId 输出引脚。理由：唯一可能的失败态是"数组维度与循环上界
 *   不一致"，而该风险已由编译期定长数组 ARRAY[0..15] 与 VAR CONSTANT
 *   DL_PACK_BIT_COUNT 双重约束消除，函数不存在任何运行期失败路径。引入一个恒为 0
 *   的错误码引脚只会增加调用方噪音。此为对"错误统一经 uErrorId 输出"规则的
 *   显式豁免，依据 ROUND_PLAN §2.6 决策记录（P3），已在手册与演进日志备案。
 *   This function intentionally has no uErrorId output: the only conceivable failure
 *   mode (array dimension vs loop bound mismatch) is removed at compile time by the
 *   fixed-size array plus a VAR CONSTANT bound, leaving no runtime failure path.
 *
 * 红线自检 (Redline)    : R1 ✓ 零全局变量表与外部变量引用 ｜ R2 ✓ 零物理 IO 地址直写
 *                         R3 ✓ 纯 IEC 61131-3（无厂商位写方言）｜ R4 ✓ 维度硬绑定 + 下标双检
 *                         R5 ✓ 全变量中英双语同行注释 ｜ R6 N/A（无状态机）｜ R7 N/A（无实例调用）
 *                         豁免项：uErrorId（见上，编译期无失败路径）
 * 修订历史 (Revision)   :
 *   2026-11-14  v1.0.0  首版入库（Phase 1 冷启动 · Level 0 批次）
 *============================================================================*)
FUNCTION FC_DL_PackBitsToWord : WORD
VAR_INPUT
    abBits     : ARRAY[0..15] OF BOOL;   // 16 路离散状态，索引 0 对应 bit0 / 16 discrete states, index 0 maps to bit0
    bInvertAll : BOOL := FALSE;          // 整体取反，适配低电平有效的报警点 / Invert all bits for active-low alarm points
END_VAR
VAR
    uResult : WORD;    // 打包结果 / Packed result word
    nIndex  : INT;     // 循环索引，值域 0..15 / Loop index, range 0..15
    uWork   : UDINT;   // 打包中间寄存器，避免 WORD 移位溢出 / Intermediate register in UDINT to avoid WORD shift overflow
END_VAR
VAR CONSTANT
    DL_PACK_BIT_COUNT : INT := 16;   // 打包位数，必须与数组维度严格一致 / Packed bit count, must equal the array dimension
END_VAR

(*------------------------------------------------------------------------------
 * 段 1｜初始化：结果清零，中间寄存器清零（不依赖实例残留值）
 *      Initialization: clear result and intermediate register
 *-----------------------------------------------------------------------------*)
uResult := 16#0000;
uWork   := 16#0000_0000;

(*------------------------------------------------------------------------------
 * 段 2｜逐位组装（边界 B1/B3）：循环上界走常量，禁止魔法数 15
 *      Bit-by-bit assembly: the loop bound comes from a constant, no magic number
 *      位序唯一约定：索引 i 的数据写入 bit i，即索引 0 → LSB
 *      Single bit-order convention: data at index i goes to bit i, index 0 = LSB
 *-----------------------------------------------------------------------------*)
FOR nIndex := 0 TO (DL_PACK_BIT_COUNT - 1) DO
    (* 数组下标上下界双检（红线 R4）：下界 0、上界 DL_PACK_BIT_COUNT-1 *)
    (* Array index double check: lower bound 0 and upper bound DL_PACK_BIT_COUNT-1 *)
    IF (nIndex >= 0) AND (nIndex <= (DL_PACK_BIT_COUNT - 1)) THEN
        IF abBits[nIndex] THEN
            (* SHL 在 UDINT 域执行，纯 IEC 语义，无厂商位写方言 *)
            (* SHL runs in the UDINT domain, pure IEC semantics, no bit-write dialect *)
            uWork := uWork OR SHL(UDINT#1, INT_TO_UDINT(nIndex));
        END_IF
    END_IF
END_FOR;

(*------------------------------------------------------------------------------
 * 段 3｜截断到 WORD 域：只保留低 16 位
 *      Truncate to the WORD domain: keep the low 16 bits only
 *-----------------------------------------------------------------------------*)
uResult := UDINT_TO_WORD(uWork);

(*------------------------------------------------------------------------------
 * 段 4｜整体取反（边界 B4）：在组装完成后一次性执行，语义清晰且少 16 次分支
 *      Global inversion executed once after assembly, clearer and cheaper
 *-----------------------------------------------------------------------------*)
IF bInvertAll THEN
    uResult := NOT uResult;
END_IF

(*------------------------------------------------------------------------------
 * 段 5｜结果回写：调用方须显式初始化 BOOL 数组，不得依赖平台默认 FALSE（边界 B5）
 *      Result write-back: callers must initialize the BOOL array explicitly
 *-----------------------------------------------------------------------------*)
FC_DL_PackBitsToWord := uResult;
END_FUNCTION

(* ---- FC_DL_ParityEvenByte.st ---- *)
(*==============================================================================
 * 组件名称 : FC_DL_ParityEvenByte ｜ 子库 : DL_Base ｜ v1.0.0 ｜ 2026-11-23
 * 平台     : CODESYS 3.5 / TwinCAT 3 / InoProShop / Machine Expert（纯 IEC，无厂商库）
 * 功能简介 : 计算字节的偶校验位：字节中 1 的个数为偶数返回 TRUE。
 *            移位 + 异或折叠 WHILE 循环实现（错位 4→2→1），不使用任何
 *            校验库函数。折叠性质：x XOR (x >> k) 不改变 1 计数的奇偶性，
 *            三轮折叠后全部 8 位信息集中到位 0。
 * 契约     : 返回 TRUE = 1 计数为偶（含全 0 字节）；输入 byVal 任意字节；
 *            纯函数无状态、同输入同输出。
 * 依赖     : 无 DL_ 内部依赖（本批自足实现）
 * 红线自检 : R1 零全局 R2 零%I/%Q R3 纯IEC R4 循环有界（错位每轮减半必归 0）
 *            R5 双语注释 R6 N/A（无状态机） R7 N/A（无定时器实例）
 * 修订历史 : 2026-11-23 R78-B1 奇偶校验族模板派生首版
 *============================================================================*)
FUNCTION FC_DL_ParityEvenByte : BOOL
VAR_INPUT
    byVal : BYTE;       // 待校验字节 / Byte to be parity-checked
END_VAR
VAR
    uX : BYTE;          // 异或折叠工作副本 / XOR-fold working copy
    nShift : INT;       // 当前错位量（4→2→1） / Current fold shift (4→2→1)
END_VAR
uX := byVal;                        // 取工作副本 / Take working copy
nShift := 4;                        // 初错位 = 半字宽 / Initial shift = half width
WHILE nShift >= 1 DO                // 折叠循环，错位每轮减半必归 0 / Fold loop, shift halves each round
    uX := uX XOR SHR(uX, nShift);   // 错位异或，奇偶性保持 / XOR fold preserves ones-parity
    nShift := nShift / 2;           // 错位减半（整除截断）/ Halve the shift
END_WHILE
FC_DL_ParityEvenByte := (uX AND 16#01) = 16#00;     // 位 0 = 全字节 1 计数奇偶 / Bit0 = parity of ones count
END_FUNCTION

(* ---- FC_DL_ParityEvenLword.st ---- *)
(*==============================================================================
 * 组件名称 : FC_DL_ParityEvenLword ｜ 子库 : DL_Base ｜ v1.0.0 ｜ 2026-11-23
 * 平台     : CODESYS 3.5 / TwinCAT 3 / InoProShop / Machine Expert（纯 IEC，无厂商库）
 * 功能简介 : 计算双字（32 位 DWORD 口径）的偶校验位：1 的个数为偶数返回
 *            TRUE。移位 + 异或折叠 WHILE 循环实现（错位 16→8→4→2→1），
 *            不使用任何校验库函数。字节/字族同算法扩位版。
 * 契约     : 返回 TRUE = 1 计数为偶（含全 0 双字）；输入 dwVal 任意双字；
 *            纯函数无状态、同输入同输出。
 * 依赖     : 无 DL_ 内部依赖（本批自足实现）
 * 红线自检 : R1 零全局 R2 零%I/%Q R3 纯IEC R4 循环有界（错位每轮减半必归 0）
 *            R5 双语注释 R6 N/A（无状态机） R7 N/A（无定时器实例）
 * 修订历史 : 2026-11-23 R78-B1 奇偶校验族模板派生首版
 *============================================================================*)
FUNCTION FC_DL_ParityEvenLword : BOOL
VAR_INPUT
    dwVal : DWORD;      // 待校验双字（32 位 DWORD） / 32-bit double word to be parity-checked
END_VAR
VAR
    uX : DWORD;         // 异或折叠工作副本 / XOR-fold working copy
    nShift : INT;       // 当前错位量（16→8→4→2→1） / Current fold shift (16→8→4→2→1)
END_VAR
uX := dwVal;                        // 取工作副本 / Take working copy
nShift := 16;                       // 初错位 = 半字宽 / Initial shift = half width
WHILE nShift >= 1 DO                // 折叠循环，错位每轮减半必归 0 / Fold loop, shift halves each round
    uX := uX XOR SHR(uX, nShift);   // 错位异或，奇偶性保持 / XOR fold preserves ones-parity
    nShift := nShift / 2;           // 错位减半（整除截断）/ Halve the shift
END_WHILE
FC_DL_ParityEvenLword := (uX AND 16#0000_0001) = 16#0000_0000;      // 位 0 = 全双字 1 计数奇偶 / Bit0 = parity of ones count
END_FUNCTION

(* ---- FC_DL_ParityEvenWord.st ---- *)
(*==============================================================================
 * 组件名称 : FC_DL_ParityEvenWord ｜ 子库 : DL_Base ｜ v1.0.0 ｜ 2026-11-23
 * 平台     : CODESYS 3.5 / TwinCAT 3 / InoProShop / Machine Expert（纯 IEC，无厂商库）
 * 功能简介 : 计算 16 位字的偶校验位：字中 1 的个数为偶数返回 TRUE。
 *            移位 + 异或折叠 WHILE 循环实现（错位 8→4→2→1），不使用
 *            任何校验库函数。字节族同算法扩位版。
 * 契约     : 返回 TRUE = 1 计数为偶（含全 0 字）；输入 wVal 任意字；
 *            纯函数无状态、同输入同输出。
 * 依赖     : 无 DL_ 内部依赖（本批自足实现）
 * 红线自检 : R1 零全局 R2 零%I/%Q R3 纯IEC R4 循环有界（错位每轮减半必归 0）
 *            R5 双语注释 R6 N/A（无状态机） R7 N/A（无定时器实例）
 * 修订历史 : 2026-11-23 R78-B1 奇偶校验族模板派生首版
 *============================================================================*)
FUNCTION FC_DL_ParityEvenWord : BOOL
VAR_INPUT
    wVal : WORD;        // 待校验 16 位字 / 16-bit word to be parity-checked
END_VAR
VAR
    uX : WORD;          // 异或折叠工作副本 / XOR-fold working copy
    nShift : INT;       // 当前错位量（8→4→2→1） / Current fold shift (8→4→2→1)
END_VAR
uX := wVal;                         // 取工作副本 / Take working copy
nShift := 8;                        // 初错位 = 半字宽 / Initial shift = half width
WHILE nShift >= 1 DO                // 折叠循环，错位每轮减半必归 0 / Fold loop, shift halves each round
    uX := uX XOR SHR(uX, nShift);   // 错位异或，奇偶性保持 / XOR fold preserves ones-parity
    nShift := nShift / 2;           // 错位减半（整除截断）/ Halve the shift
END_WHILE
FC_DL_ParityEvenWord := (uX AND 16#0001) = 16#0000;     // 位 0 = 全字 1 计数奇偶 / Bit0 = parity of ones count
END_FUNCTION

(* ---- FC_DL_ParityOddByte.st ---- *)
(*==============================================================================
 * 组件名称 : FC_DL_ParityOddByte ｜ 子库 : DL_Base ｜ v1.0.0 ｜ 2026-11-23
 * 平台     : CODESYS 3.5 / TwinCAT 3 / InoProShop / Machine Expert（纯 IEC，无厂商库）
 * 功能简介 : 计算字节的奇校验位：字节中 1 的个数为奇数返回 TRUE。
 *            移位 + 异或折叠 WHILE 循环实现（错位 4→2→1），不使用任何
 *            校验库函数。与偶校验件同族同算法，仅判定取反。
 * 契约     : 返回 TRUE = 1 计数为奇；输入 byVal 任意字节（全 0 返回 FALSE）；
 *            纯函数无状态、同输入同输出。
 * 依赖     : 无 DL_ 内部依赖（本批自足实现）
 * 红线自检 : R1 零全局 R2 零%I/%Q R3 纯IEC R4 循环有界（错位每轮减半必归 0）
 *            R5 双语注释 R6 N/A（无状态机） R7 N/A（无定时器实例）
 * 修订历史 : 2026-11-23 R78-B1 奇偶校验族模板派生首版
 *============================================================================*)
FUNCTION FC_DL_ParityOddByte : BOOL
VAR_INPUT
    byVal : BYTE;       // 待校验字节 / Byte to be parity-checked
END_VAR
VAR
    uX : BYTE;          // 异或折叠工作副本 / XOR-fold working copy
    nShift : INT;       // 当前错位量（4→2→1） / Current fold shift (4→2→1)
END_VAR
uX := byVal;                        // 取工作副本 / Take working copy
nShift := 4;                        // 初错位 = 半字宽 / Initial shift = half width
WHILE nShift >= 1 DO                // 折叠循环，错位每轮减半必归 0 / Fold loop, shift halves each round
    uX := uX XOR SHR(uX, nShift);   // 错位异或，奇偶性保持 / XOR fold preserves ones-parity
    nShift := nShift / 2;           // 错位减半（整除截断）/ Halve the shift
END_WHILE
FC_DL_ParityOddByte := (uX AND 16#01) = 16#01;      // 位 0 = 1 计数奇偶，奇返回 TRUE / Bit0 = parity, TRUE if odd
END_FUNCTION

(* ---- FC_DL_ParityOddLword.st ---- *)
(*==============================================================================
 * 组件名称 : FC_DL_ParityOddLword ｜ 子库 : DL_Base ｜ v1.0.0 ｜ 2026-11-23
 * 平台     : CODESYS 3.5 / TwinCAT 3 / InoProShop / Machine Expert（纯 IEC，无厂商库）
 * 功能简介 : 计算双字（32 位 DWORD 口径）的奇校验位：1 的个数为奇数返回
 *            TRUE。移位 + 异或折叠 WHILE 循环实现（错位 16→8→4→2→1），
 *            不使用任何校验库函数。与偶校验件同族同算法，仅判定取反。
 * 契约     : 返回 TRUE = 1 计数为奇；输入 dwVal 任意双字（全 0 返回 FALSE）；
 *            纯函数无状态、同输入同输出。
 * 依赖     : 无 DL_ 内部依赖（本批自足实现）
 * 红线自检 : R1 零全局 R2 零%I/%Q R3 纯IEC R4 循环有界（错位每轮减半必归 0）
 *            R5 双语注释 R6 N/A（无状态机） R7 N/A（无定时器实例）
 * 修订历史 : 2026-11-23 R78-B1 奇偶校验族模板派生首版
 *============================================================================*)
FUNCTION FC_DL_ParityOddLword : BOOL
VAR_INPUT
    dwVal : DWORD;      // 待校验双字（32 位 DWORD） / 32-bit double word to be parity-checked
END_VAR
VAR
    uX : DWORD;         // 异或折叠工作副本 / XOR-fold working copy
    nShift : INT;       // 当前错位量（16→8→4→2→1） / Current fold shift (16→8→4→2→1)
END_VAR
uX := dwVal;                        // 取工作副本 / Take working copy
nShift := 16;                       // 初错位 = 半字宽 / Initial shift = half width
WHILE nShift >= 1 DO                // 折叠循环，错位每轮减半必归 0 / Fold loop, shift halves each round
    uX := uX XOR SHR(uX, nShift);   // 错位异或，奇偶性保持 / XOR fold preserves ones-parity
    nShift := nShift / 2;           // 错位减半（整除截断）/ Halve the shift
END_WHILE
FC_DL_ParityOddLword := (uX AND 16#0000_0001) = 16#0000_0001;       // 位 0 = 1 计数奇偶，奇返回 TRUE / Bit0 = parity, TRUE if odd
END_FUNCTION

(* ---- FC_DL_ParityOddWord.st ---- *)
(*==============================================================================
 * 组件名称 : FC_DL_ParityOddWord ｜ 子库 : DL_Base ｜ v1.0.0 ｜ 2026-11-23
 * 平台     : CODESYS 3.5 / TwinCAT 3 / InoProShop / Machine Expert（纯 IEC，无厂商库）
 * 功能简介 : 计算 16 位字的奇校验位：字中 1 的个数为奇数返回 TRUE。
 *            移位 + 异或折叠 WHILE 循环实现（错位 8→4→2→1），不使用
 *            任何校验库函数。与偶校验件同族同算法，仅判定取反。
 * 契约     : 返回 TRUE = 1 计数为奇；输入 wVal 任意字（全 0 返回 FALSE）；
 *            纯函数无状态、同输入同输出。
 * 依赖     : 无 DL_ 内部依赖（本批自足实现）
 * 红线自检 : R1 零全局 R2 零%I/%Q R3 纯IEC R4 循环有界（错位每轮减半必归 0）
 *            R5 双语注释 R6 N/A（无状态机） R7 N/A（无定时器实例）
 * 修订历史 : 2026-11-23 R78-B1 奇偶校验族模板派生首版
 *============================================================================*)
FUNCTION FC_DL_ParityOddWord : BOOL
VAR_INPUT
    wVal : WORD;        // 待校验 16 位字 / 16-bit word to be parity-checked
END_VAR
VAR
    uX : WORD;          // 异或折叠工作副本 / XOR-fold working copy
    nShift : INT;       // 当前错位量（8→4→2→1） / Current fold shift (8→4→2→1)
END_VAR
uX := wVal;                         // 取工作副本 / Take working copy
nShift := 8;                        // 初错位 = 半字宽 / Initial shift = half width
WHILE nShift >= 1 DO                // 折叠循环，错位每轮减半必归 0 / Fold loop, shift halves each round
    uX := uX XOR SHR(uX, nShift);   // 错位异或，奇偶性保持 / XOR fold preserves ones-parity
    nShift := nShift / 2;           // 错位减半（整除截断）/ Halve the shift
END_WHILE
FC_DL_ParityOddWord := (uX AND 16#0001) = 16#0001;      // 位 0 = 1 计数奇偶，奇返回 TRUE / Bit0 = parity, TRUE if odd
END_FUNCTION

(* ---- FC_DL_PipeInsulationLossCalc.st ---- *)
(*
  Component : FC_DL_PipeInsulationLossCalc
  Category  : DL_Base
  Function  : 圆筒管道保温散热 q = 2πλ(Ti−To)/ln(r2/r1)，单位 W/m
  Complexity: C2
  开源溯源 : DLF 内部原创（R94 族模板派生）；参考语义来源见 SOURCE_HUNTING_MATRIX.md
  规则遵从 : R1-R16
  契约     : 输入 rTiC 管内介质温度 [℃]、rToC 环境温度 [℃]、rLambdaWmK 保温材料导热系数 [W/(m·K)]、
             rInnerDiaMm 管道外径（保温内径） [mm]、rThickMm 保温层厚度 [mm]；
             输出 rQwm 单位管长热损 [W/m]、rQTotalW 给定管长总热损 [W]、rOuterDiaMm 保温外径 [mm]、
             xValid 有效标志、nFaultCode 故障码。
  边界     : 半径比 r2/r1 为无量纲量，故内外径可用 [mm] 直接参与对数（无需折米）；
             r1 须 >1.0E-6 [mm]、r2 须 > r1（厚度 >0）；ln(r2/r1) 须 >1.0E-9；
             导热系数须 >0；管长 rLengthM 用于总热损，为 0 时总热损输出 0（不判故障）。
  码位     : 9801 输入非有限（故障级）；9802 半径比或导热系数越域（故障级）。
*)
FUNCTION FC_DL_PipeInsulationLossCalc : BOOL
VAR_INPUT
    rTiC        : LREAL := 150.0;     // 管内介质温度 [℃] EN: the medium temperature inside the pipe
    rToC        : LREAL := 25.0;      // 环境温度 [℃] EN: the ambient temperature
    rLambdaWmK  : LREAL := 0.045;     // 保温材料导热系数 [W/(m·K)] EN: the thermal conductivity of the insulation
    rInnerDiaMm : LREAL := 108.0;     // 管道外径即保温内径 [mm] EN: the pipe outer diameter acting as the insulation inner diameter
    rThickMm    : LREAL := 50.0;      // 保温层厚度 [mm] EN: the insulation thickness
    rLengthM    : LREAL := 10.0;      // 参与总热损的管长 [m] EN: the pipe length used for the total loss
END_VAR
VAR_OUTPUT
    rQwm       : LREAL;               // 单位管长热损 [W/m] EN: the heat loss per metre of pipe
    rQTotalW   : LREAL;               // 管长总热损 [W] EN: the total heat loss over the given length
    rOuterDiaMm: LREAL;               // 保温外径 [mm] EN: the insulation outer diameter
    xValid     : BOOL;                // 输出可信标志 EN: the outputs are valid
    nFaultCode : INT;                 // 0=无故障 9801=输入非有限 9802=半径比或导热系数越域 EN: zero none, 9801 non finite, 9802 radius ratio or conductivity out of range
END_VAR
VAR
    xFinAll : BOOL;                   // 六个浮点入参有限 EN: all six floating inputs are finite
    rR1     : LREAL;                  // 保温内半径 [mm] EN: the insulation inner radius
    rR2     : LREAL;                  // 保温外半径 [mm] EN: the insulation outer radius
    rRat    : LREAL;                  // 半径比 r2/r1 [-] EN: the radius ratio
    rLn     : LREAL;                  // 半径比对数 [-] EN: the logarithm of the radius ratio
    rQ      : LREAL;                  // 单位热损中间值 [W/m] EN: the interim loss per metre
END_VAR
VAR CONSTANT
    DL_PIL_Z       : LREAL := 0.0;                  // 浮点零常量 EN: the floating point zero constant
    DL_PIL_TWO     : LREAL := 2.0;                  // 直径转半径系数 EN: the diameter to radius factor
    DL_PIL_PI2     : LREAL := 6.2831853071795865;   // 2π（LREAL 精度） [-] EN: twice the circle ratio at LREAL precision
    DL_PIL_MIN     : LREAL := 1.0E-9;               // 对数与半径的下限 EN: the lower bound of the logarithm and the radius
    DL_PIL_C_BAD   : INT := 9801;                   // 输入非有限 EN: a non finite input
    DL_PIL_C_RANGE : INT := 9802;                   // 半径比或导热系数越域 EN: the radius ratio or the conductivity is out of range
END_VAR

// 段1｜出口预置
FC_DL_PipeInsulationLossCalc := FALSE;   // 返回值预置假 EN: preset the return value to false
rQwm := DL_PIL_Z;                        // 单位热损预置零 [W/m] EN: preset the loss per metre to zero
rQTotalW := DL_PIL_Z;                    // 总热损预置零 [W] EN: preset the total loss to zero
rOuterDiaMm := DL_PIL_Z;                 // 外径预置零 [mm] EN: preset the outer diameter to zero
xValid := FALSE;                         // 有效标志预置假 EN: preset the validity flag to false
nFaultCode := 0;                         // 故障码预置零 EN: preset the fault code to zero

// 段2｜非有限闸：六输入全列
xFinAll := (rTiC = rTiC) AND ((rTiC - rTiC) = DL_PIL_Z)
        AND (rToC = rToC) AND ((rToC - rToC) = DL_PIL_Z)
        AND (rLambdaWmK = rLambdaWmK) AND ((rLambdaWmK - rLambdaWmK) = DL_PIL_Z)
        AND (rInnerDiaMm = rInnerDiaMm) AND ((rInnerDiaMm - rInnerDiaMm) = DL_PIL_Z)
        AND (rThickMm = rThickMm) AND ((rThickMm - rThickMm) = DL_PIL_Z)
        AND (rLengthM = rLengthM) AND ((rLengthM - rLengthM) = DL_PIL_Z);   // 六输入有限性 EN: the finiteness of all six inputs
IF NOT xFinAll THEN                                                          // 非有限出口 EN: leave early on a non finite input
    nFaultCode := DL_PIL_C_BAD;                                              // 非有限码 EN: the non finite code
    RETURN;                                                                  // 早退 EN: return early
END_IF

// 段3｜域闸：内半径为分母须够大、厚度为正、导热系数为正、管长非负
rR1 := rInnerDiaMm / DL_PIL_TWO;                                             // 保温内半径 [mm] EN: the insulation inner radius
rR2 := rR1 + rThickMm;                                                       // 保温外半径 [mm] EN: the insulation outer radius
rOuterDiaMm := rInnerDiaMm + DL_PIL_TWO * rThickMm;                          // 保温外径 [mm] EN: the insulation outer diameter
IF (rR1 < DL_PIL_MIN) OR (rThickMm <= DL_PIL_Z) OR (rLambdaWmK <= DL_PIL_Z) OR (rLengthM < DL_PIL_Z) THEN
    nFaultCode := DL_PIL_C_RANGE;                                            // 越域码 EN: the out of range code
    RETURN;                                                                  // 早退 EN: return early
END_IF

// 段4｜主体：q = 2πλΔT / ln(r2/r1)
rRat := rR2 / rR1;                                                           // 半径比，分母已过下限 [-] EN: the radius ratio, the divisor passed the gate
rLn := LN(rRat);                                                             // 半径比对数 [-] EN: the logarithm of the radius ratio
IF ABS(rLn) < DL_PIL_MIN THEN                                                // 对数下限（厚度趋零） EN: the logarithm gate for a vanishing thickness
    nFaultCode := DL_PIL_C_RANGE;                                            // 越域码 EN: the out of range code
    RETURN;                                                                  // 早退 EN: return early
END_IF
rQ := (DL_PIL_PI2 * rLambdaWmK * (rTiC - rToC)) / rLn;                        // 单位管长热损，正负随温差 [W/m] EN: the loss per metre carrying the temperature difference sign

// 段5｜结果复检与出口
IF rQ <> rQ THEN                                                             // 复检：非有限 EN: recheck for a non finite value
    nFaultCode := DL_PIL_C_RANGE;                                            // 复检失败码 EN: the recheck failure code
    RETURN;                                                                  // 早退，出口保持零哨兵 EN: return early with the zero sentinels
END_IF
rQwm := rQ;                                                                  // 单位热损出口 [W/m] EN: the loss per metre output
rQTotalW := rQ * rLengthM;                                                   // 总热损 = 单位热损 × 管长 [W] EN: the total loss over the length
xValid := TRUE;                                                              // 结果可信 EN: the results are valid
FC_DL_PipeInsulationLossCalc := TRUE;                                         // 返回真 EN: return true
END_FUNCTION

(* ---- FC_DL_PriorityEncodeWord.st ---- *)
(*
  Name        : FC_DL_PriorityEncodeWord
  Category    : DL_Base
  Version     : 1.0.0
  Purpose     : 位串优先编码：返回最高或最低置 1 位的位序号（1..32），无置位返回 0 号哨兵；/ Priority encoding: return the bit number (1..32) of the highest or lowest set bit, sentinel 0 when none
  溯源        : 借 t2-1-lgf·bitlogic 的分类/参数域组织，clean-room 实现
  Boundary    : ① 位序号口径为 1 基（1..32），哨兵 0 表示「无置位」，二者不重叠；
                ② 移位量恒 0..31 < 32，禁 SHL(x, 位宽)；
                ③ 结果上限 32 钳位（防下游数组下标越界，R308）；
                ④ 纯位运算无除零；整型入参无 NaN 路径。
*)
FUNCTION FC_DL_PriorityEncodeWord : INT
VAR_INPUT
    dwBits   : DWORD := 0;                   (* 待编码位串（32 位解释）[-] / Bit string to encode, 32-bit *)
    xHighest : BOOL := TRUE;                 (* TRUE = 最高置位优先；FALSE = 最低置位优先 [-] / Highest-set or lowest-set priority *)
END_VAR
VAR
    nIdx   : INT;                            (* 位序号游标 0..31（FOR 自复位，R227）[-] / Bit index cursor 0..31 *)
    nFound : INT;                            (* 命中位号 1..32；0 = 无置位哨兵 [-] / Hit bit number 1..32, 0 = none *)
    dwMask : DWORD;                          (* 单热掩码，初值 1 后逐位左移 [-] / Walking-one mask *)
END_VAR
VAR CONSTANT
    DL_PEW_WIDTH : INT   := 32;              (* DWORD 位宽（移位量上界基准）[位] / DWORD bit width *)
    DL_PEW_NONE  : INT   := 0;               (* 无置位哨兵位号（与 1..32 不重叠）[-] / No-bit sentinel *)
    DL_PEW_ONE   : DWORD := 1;               (* 单热掩码初值 [-] / Initial mask *)
    DL_PEW_ZERO  : DWORD := 0;               (* 位串零常量 [-] / Zero constant *)
END_VAR

(* —— 段 1：单拍量预清零（每拍全路径派生，R107） —— *)
nFound := DL_PEW_NONE;                       (* 哨兵预置：仅命中分支改写 / Sentinel preset *)
dwMask := DL_PEW_ONE;                        (* 掩码从最低位起扫 / Mask starts at LSB *)

(* —— 段 2：逐位扫描（单循环 + 优先级策略，两口径同一遍历） —— *)
FOR nIdx := 0 TO DL_PEW_WIDTH - 1 DO
    IF (dwBits AND dwMask) <> DL_PEW_ZERO THEN
        IF xHighest THEN
            nFound := nIdx + 1;              (* 最高优先：持续覆盖，末次命中即最高位 / Highest: last hit wins *)
        ELSIF nFound = DL_PEW_NONE THEN
            nFound := nIdx + 1;              (* 最低优先：首个命中即锁定，后续不覆盖 / Lowest: first hit locks *)
        END_IF
    END_IF
    dwMask := SHL(dwMask, 1);                (* 掩码左移（1..31 < 32，无越界） / Shift mask, amount < width *)
END_FOR

(* —— 段 3：输出上限钳位（1..32 或哨兵 0，二者互斥且均在合法域） —— *)
IF nFound > DL_PEW_WIDTH THEN
    nFound := DL_PEW_WIDTH;                  (* 上限饱和 32：理论不可达，防御性 / Upper saturation, defensive *)
ELSIF nFound < DL_PEW_NONE THEN
    nFound := DL_PEW_NONE;                   (* 下限兜底到哨兵 / Lower fallback to sentinel *)
END_IF
FC_DL_PriorityEncodeWord := nFound;          (* 返回位号或哨兵 0 / Return bit number or sentinel 0 *)
END_FUNCTION

(* ---- FC_DL_Q15AbsSat.st ---- *)
(*
  FC_DL_Q15AbsSat —— Q15 取绝对值饱和，正确处理 -32768 边界
  分类：DL_Base | 复杂度：1 | 轮次：R86
  开源溯源：道莅原创（clean-room 自研，纯 IEC 61131-3 通用算法），无外部代码引用
  许可证：MIT
  职责：Q15 取绝对值；-32768 的绝对值 32768 超出 Q15 上界，饱和回 32767 并置 xSat。
  契约：iIn 输入 [Q15]；返回绝对值 [Q15]；xSat 报告 -32768 边界饱和（信息级）。
  边界：不走 ABS(INT)（-32768 上溢），先升 DINT 再取绝对值；零全局、零物理地址、零库件依赖。
*)
FUNCTION FC_DL_Q15AbsSat : INT
VAR_INPUT
    iIn : INT := 0;                   // 输入操作数 [Q15] / The input operand in Q15
END_VAR
VAR_OUTPUT
    xSat : BOOL;                      // 边界饱和标志（信息级） [—] / The boundary saturation flag
END_VAR
VAR
    diAbs : DINT;                     // 双字绝对值暂存 [Q15] / The double word absolute stage
END_VAR
VAR CONSTANT
    Q15_MAX : DINT := 32767;          // Q15 上界 [-] / The Q15 upper bound
END_VAR

xSat := FALSE;                                        // 饱和标志预置假 / preset the saturation flag false
diAbs := ABS(INT_TO_DINT(iIn));                       // 升 DINT 后取绝对值（-32768 在 DINT 域安全） [Q15] / absolute in DINT
IF diAbs > Q15_MAX THEN                               // 仅 -32768 会命中此分支 / only minus 32768 hits this branch
    FC_DL_Q15AbsSat := DINT_TO_INT(Q15_MAX);          // 饱和到 Q15_MAX [Q15] / saturate high
    xSat := TRUE;                                     // 置饱和标志 [—] / raise the saturation flag
ELSE
    FC_DL_Q15AbsSat := DINT_TO_INT(diAbs);            // 界内直接转换 [Q15] / in range conversion
END_IF
END_FUNCTION

(* ---- FC_DL_Q15AddSat.st ---- *)
(*
  FC_DL_Q15AddSat —— Q15 定点加法饱和，越界钳到 Q15_MAX/Q15_MIN
  分类：DL_Base | 复杂度：2 | 轮次：R86
  开源溯源：道莅原创（clean-room 自研，纯 IEC 61131-3 通用算法），无外部代码引用
  许可证：MIT
  职责：Q15 域两数相加，中间用 DINT 承载，结果按 Q15 上下界饱和。
  契约：输入 iA / iB 为 Q15 操作数；返回 Q15 和；xSat 报告本拍发生饱和（信息级）。
  边界：DINT 中间量 + 上下界双判，无除法、无浮点比较；零全局、零物理地址、零库件依赖。
*)
FUNCTION FC_DL_Q15AddSat : INT
VAR_INPUT
    iA : INT := 0;                    // 加数 A [Q15] / The addend A in Q15
    iB : INT := 0;                    // 加数 B [Q15] / The addend B in Q15
END_VAR
VAR_OUTPUT
    xSat : BOOL;                      // 饱和发生标志（信息级） [—] / The saturation flag, informational
END_VAR
VAR
    diSum : DINT;                     // 双字中间和 [Q15] / The double word intermediate sum
END_VAR
VAR CONSTANT
    Q15_MAX : DINT := 32767;          // Q15 上界 [-] / The Q15 upper bound
    Q15_MIN : DINT := -32768;         // Q15 下界 [-] / The Q15 lower bound
END_VAR

xSat := FALSE;                                        // 饱和标志预置假 / preset the saturation flag false
diSum := INT_TO_DINT(iA) + INT_TO_DINT(iB);           // 双字域求和（|和| <= 65535 不溢出） [Q15] / sum in DINT
IF diSum > Q15_MAX THEN                               // 上越界 / above the upper bound
    FC_DL_Q15AddSat := DINT_TO_INT(Q15_MAX);          // 饱和到 Q15_MAX [Q15] / saturate high
    xSat := TRUE;                                     // 置饱和标志 [—] / raise the saturation flag
ELSIF diSum < Q15_MIN THEN                            // 下越界 / below the lower bound
    FC_DL_Q15AddSat := DINT_TO_INT(Q15_MIN);          // 饱和到 Q15_MIN [Q15] / saturate low
    xSat := TRUE;                                     // 置饱和标志 [—] / raise the saturation flag
ELSE
    FC_DL_Q15AddSat := DINT_TO_INT(diSum);            // 界内直接转换 [Q15] / in range conversion
END_IF
END_FUNCTION

(* ---- FC_DL_Q15DivSafe.st ---- *)
(*
  FC_DL_Q15DivSafe —— Q15 安全除法，除零与商越界双保护
  分类：DL_Base | 复杂度：2 | 轮次：R86
  开源溯源：道莅原创（clean-room 自研，纯 IEC 61131-3 通用算法），无外部代码引用
  许可证：MIT
  职责：Q15 除以 Q15 得 Q15：先把被除数放大 32768 倍（DINT 界内），再整除并按 Q15 饱和。
  契约：iNum 被除数 [Q15]、iDen 除数 [Q15]；返回商 [Q15]；xValid 除数为零时为 FALSE（商给零哨兵）。
  边界：① 除零前置判（R4）；② 商越界双侧饱和；③ 被除数放大后 |值| <= 1.074e9 已证不溢出；
        ④ 零全局、零物理地址、零库件依赖。
*)
FUNCTION FC_DL_Q15DivSafe : INT
VAR_INPUT
    iNum : INT := 0;                  // 被除数 [Q15] / The dividend in Q15
    iDen : INT := 0;                  // 除数 [Q15] / The divisor in Q15
END_VAR
VAR_OUTPUT
    xValid : BOOL;                    // 商可信（除数非零） [—] / The quotient is valid when the divisor is non zero
    xSat   : BOOL;                    // 商越界饱和标志（信息级） [—] / The quotient saturation flag
END_VAR
VAR
    diNum : DINT;                     // 放大后的被除数 [Q30] / The scaled dividend in Q30
    diQ   : DINT;                     // 商暂存 [Q15] / The quotient stage
END_VAR
VAR CONSTANT
    Q15_MAX  : DINT := 32767;         // Q15 上界 [-] / The Q15 upper bound
    Q15_MIN  : DINT := -32768;        // Q15 下界 [-] / The Q15 lower bound
    DL_QD_SC : DINT := 32768;         // 定标因子（2^15） [-] / The Q15 scaling factor
    DL_QD_Z  : DINT := 0;             // 整型零常量 [-] / The integer zero constant
END_VAR

xValid := FALSE;                                      // 可信位预置假 / preset the valid flag false
xSat := FALSE;                                        // 饱和标志预置假 / preset the saturation flag false
IF iDen = DL_QD_Z THEN                                // 除数为零（除零防护，前置判） / the divisor is zero
    FC_DL_Q15DivSafe := DINT_TO_INT(DL_QD_Z);         // 商给零哨兵 [Q15] / the zero sentinel quotient
ELSE
    diNum := INT_TO_DINT(iNum) * DL_QD_SC;            // 被除数放大 15 位（|值| <= 1.074e9 界内） [Q30] / scale the dividend
    diQ := diNum / INT_TO_DINT(iDen);                 // 整除得商（分母已证非零） [Q15] / integer division
    IF diQ > Q15_MAX THEN                             // 商上越界 / the quotient above the upper bound
        FC_DL_Q15DivSafe := DINT_TO_INT(Q15_MAX);     // 饱和到 Q15_MAX [Q15] / saturate high
        xSat := TRUE;                                 // 置饱和标志 [—] / raise the saturation flag
    ELSIF diQ < Q15_MIN THEN                          // 商下越界 / the quotient below the lower bound
        FC_DL_Q15DivSafe := DINT_TO_INT(Q15_MIN);     // 饱和到 Q15_MIN [Q15] / saturate low
        xSat := TRUE;                                 // 置饱和标志 [—] / raise the saturation flag
    ELSE
        FC_DL_Q15DivSafe := DINT_TO_INT(diQ);         // 界内直接转换 [Q15] / in range conversion
    END_IF
    xValid := TRUE;                                   // 除法成功，商可信 [—] / the division succeeded
END_IF
END_FUNCTION

(* ---- FC_DL_Q15Lerp.st ---- *)
(*
  FC_DL_Q15Lerp —— Q15 线性插值，alpha 定点，端点饱和
  分类：DL_Base | 复杂度：2 | 轮次：R86
  开源溯源：道莅原创（clean-room 自研，纯 IEC 61131-3 通用算法），无外部代码引用
  许可证：MIT
  职责：按 Q15 权重做线性插值：out = A + (B - A) * alpha / 32767；alpha = 0 得 A，alpha = 32767 得 B。
  契约：iA 起点 [Q15]、iB 终点 [Q15]、iAlpha 权重 [Q15 归一化 0..32767]；返回插值 [Q15]；xSat 报告饱和。
  边界：① 乘积 |diD * alpha| <= 65535 * 32767 = 2.147e9 界内已证；② 除数恒为常量 32767 非零；
        ③ 端点经饱和钳位保证不越 Q15；零全局、零物理地址、零库件依赖。
*)
FUNCTION FC_DL_Q15Lerp : INT
VAR_INPUT
    iA      : INT := 0;               // 插值起点值 [Q15] / The interpolation start value in Q15
    iB      : INT := 0;               // 插值终点值 [Q15] / The interpolation end value in Q15
    iAlpha  : INT := 0;               // 归一化权重 0..32767 [Q15] / The normalised weight in Q15
END_VAR
VAR_OUTPUT
    xSat : BOOL;                      // 饱和发生标志（信息级） [—] / The saturation flag, informational
END_VAR
VAR
    diD   : DINT;                     // 端点差 [Q15] / The endpoint difference
    diP   : DINT;                     // 差乘权重（Q30 量级，界内已证） [Q30] / The scaled product
    diQ   : DINT;                     // 插值增量 [Q15] / The interpolation increment
    diR   : DINT;                     // 插值结果暂存 [Q15] / The interpolation result stage
END_VAR
VAR CONSTANT
    Q15_MAX   : DINT := 32767;        // Q15 上界 [-] / The Q15 upper bound
    Q15_MIN   : DINT := -32768;       // Q15 下界 [-] / The Q15 lower bound
    DL_QL_ONE : DINT := 32767;        // 归一化满量程（2^15 - 1） [-] / The normalisation full scale
    DL_QL_Z   : DINT := 0;            // 整型零常量 [-] / The integer zero constant
END_VAR

xSat := FALSE;                                        // 饱和标志预置假 / preset the saturation flag false
diD := INT_TO_DINT(iB) - INT_TO_DINT(iA);             // 端点差（|差| <= 65535） [Q15] / the endpoint difference
diP := diD * INT_TO_DINT(iAlpha);                     // 差乘权重（|积| <= 2.147e9 界内已证） [Q30] / the scaled product
diQ := diP / DL_QL_ONE;                               // 除以归一化满量程（常量非零） [Q15] / divide by the full scale
diR := INT_TO_DINT(iA) + diQ;                         // 起点加增量 [Q15] / the start plus the increment
IF diR > Q15_MAX THEN                                 // 上越界 / above the upper bound
    FC_DL_Q15Lerp := DINT_TO_INT(Q15_MAX);            // 饱和到 Q15_MAX [Q15] / saturate high
    xSat := TRUE;                                     // 置饱和标志 [—] / raise the saturation flag
ELSIF diR < Q15_MIN THEN                              // 下越界 / below the lower bound
    FC_DL_Q15Lerp := DINT_TO_INT(Q15_MIN);            // 饱和到 Q15_MIN [Q15] / saturate low
    xSat := TRUE;                                     // 置饱和标志 [—] / raise the saturation flag
ELSE
    FC_DL_Q15Lerp := DINT_TO_INT(diR);                // 界内直接转换 [Q15] / in range conversion
END_IF
END_FUNCTION

(* ---- FC_DL_Q15MulSat.st ---- *)
(*
  FC_DL_Q15MulSat —— Q15 乘 Q15 得 Q15，中间 DINT 防溢出，含右移舍入
  分类：DL_Base | 复杂度：2 | 轮次：R86
  开源溯源：道莅原创（clean-room 自研，纯 IEC 61131-3 通用算法），无外部代码引用
  许可证：MIT
  职责：Q15 × Q15 得 Q30（DINT 承载），加半偏置后除 32768 得 Q15，结果按 Q15 上下界饱和。
  契约：输入 iA / iB 为 Q15 操作数；返回 Q15 积；xSat 报告饱和（信息级）。
  边界：① 舍入偏置前先做「极限值反算」防 DINT 溢出；② 用乘 32768 表达定标，规避 SHL 方言差异；
        ③ 无除法风险（除数恒为常量 32768 非零）；零全局、零物理地址、零库件依赖。
*)
FUNCTION FC_DL_Q15MulSat : INT
VAR_INPUT
    iA : INT := 0;                    // 乘数 A [Q15] / The multiplier A in Q15
    iB : INT := 0;                    // 乘数 B [Q15] / The multiplier B in Q15
END_VAR
VAR_OUTPUT
    xSat : BOOL;                      // 饱和发生标志（信息级） [—] / The saturation flag, informational
END_VAR
VAR
    diProd : DINT;                    // 乘积（Q30） [Q30] / The product in Q30
    diQ : DINT;                       // 舍入右移后的 Q15 暂存 [Q15] / The rounded Q15 stage
END_VAR
VAR CONSTANT
    Q15_MAX   : DINT := 32767;        // Q15 上界 [-] / The Q15 upper bound
    Q15_MIN   : DINT := -32768;       // Q15 下界 [-] / The Q15 lower bound
    DL_QM_RND : DINT := 16384;        // 四舍五入偏置（2^14） [-] / The rounding bias
    DL_QM_SC  : DINT := 32768;        // 定标因子（2^15） [-] / The Q15 scaling factor
    DL_QM_HI  : DINT := 2147483647;   // DINT 上限（反算用） [-] / The DINT maximum
    DL_QM_LO  : DINT := -2147483647;  // DINT 下限近似（偏置在界侧相加，避下溢） [-] / The DINT minimum approximation
    DL_QM_Z   : DINT := 0;            // 整型零常量 [-] / The integer zero constant
END_VAR

xSat := FALSE;                                        // 饱和标志预置假 / preset the saturation flag false
diProd := INT_TO_DINT(iA) * INT_TO_DINT(iB);          // Q15 乘 Q15 得 Q30（|积| <= 1.074e9 界内） / Q15 times Q15
IF diProd > (DL_QM_HI - DL_QM_RND) THEN               // 加偏置前上界反算防溢出 / upper bound reverse check before rounding
    FC_DL_Q15MulSat := DINT_TO_INT(Q15_MAX);          // 直接饱和到上界 [Q15] / saturate high
    xSat := TRUE;                                     // 置饱和标志 [—] / raise the saturation flag
ELSIF diProd < (DL_QM_LO + DL_QM_RND) THEN            // 加偏置前下界反算防溢出（偏置加在界侧，避 DINT 下溢） / lower bound reverse check
    FC_DL_Q15MulSat := DINT_TO_INT(Q15_MIN);          // 直接饱和到下界 [Q15] / saturate low
    xSat := TRUE;                                     // 置饱和标志 [—] / raise the saturation flag
ELSE
    IF diProd >= DL_QM_Z THEN                         // 非负做加偏置舍入 / non negative rounding
        diQ := (diProd + DL_QM_RND) / DL_QM_SC;       // 四舍五入右移 15 位 [Q15] / rounded shift right
    ELSE
        diQ := (diProd - DL_QM_RND) / DL_QM_SC;       // 负值做减偏置舍入 [Q15] / rounded shift right
    END_IF
    IF diQ > Q15_MAX THEN                             // 上越界 / above the upper bound
        FC_DL_Q15MulSat := DINT_TO_INT(Q15_MAX);      // 饱和到 Q15_MAX [Q15] / saturate high
        xSat := TRUE;                                 // 置饱和标志 [—] / raise the saturation flag
    ELSIF diQ < Q15_MIN THEN                          // 下越界 / below the lower bound
        FC_DL_Q15MulSat := DINT_TO_INT(Q15_MIN);      // 饱和到 Q15_MIN [Q15] / saturate low
        xSat := TRUE;                                 // 置饱和标志 [—] / raise the saturation flag
    ELSE
        FC_DL_Q15MulSat := DINT_TO_INT(diQ);          // 界内直接转换 [Q15] / in range conversion
    END_IF
END_IF
END_FUNCTION

(* ---- FC_DL_Q15NegSat.st ---- *)
(*
  FC_DL_Q15NegSat —— Q15 取负饱和，-32768 不回绕
  分类：DL_Base | 复杂度：1 | 轮次：R86
  开源溯源：道莅原创（clean-room 自研，纯 IEC 61131-3 通用算法），无外部代码引用
  许可证：MIT
  职责：Q15 取负；-32768 的相反数 32768 超出 Q15 上界，饱和回 32767 并置 xSat。
  契约：iIn 输入 [Q15]；返回相反数 [Q15]；xSat 报告 -32768 边界饱和（信息级）。
  边界：不使用一元负号直接作用于 INT（-32768 回绕），先在 DINT 域取负；零全局、零物理地址、零库件依赖。
*)
FUNCTION FC_DL_Q15NegSat : INT
VAR_INPUT
    iIn : INT := 0;                   // 输入操作数 [Q15] / The input operand in Q15
END_VAR
VAR_OUTPUT
    xSat : BOOL;                      // 边界饱和标志（信息级） [—] / The boundary saturation flag
END_VAR
VAR
    diNeg : DINT;                     // 双字取负暂存 [Q15] / The double word negation stage
END_VAR
VAR CONSTANT
    Q15_MAX : DINT := 32767;          // Q15 上界 [-] / The Q15 upper bound
    Q15_MIN : DINT := -32768;         // Q15 下界 [-] / The Q15 lower bound
    DL_QN_Z : DINT := 0;              // 整型零常量 [-] / The integer zero constant
END_VAR

xSat := FALSE;                                        // 饱和标志预置假 / preset the saturation flag false
diNeg := DL_QN_Z - INT_TO_DINT(iIn);                  // 双字域取负（-32768 → 32768 在 DINT 域安全） [Q15] / negate in DINT
IF diNeg > Q15_MAX THEN                               // 仅 -32768 会命中此分支 / only minus 32768 hits this branch
    FC_DL_Q15NegSat := DINT_TO_INT(Q15_MAX);          // 饱和到 Q15_MAX [Q15] / saturate high
    xSat := TRUE;                                     // 置饱和标志 [—] / raise the saturation flag
ELSIF diNeg < Q15_MIN THEN                            // 下越界（本件数学上不可达，防御保留） / below the lower bound
    FC_DL_Q15NegSat := DINT_TO_INT(Q15_MIN);          // 饱和到 Q15_MIN [Q15] / saturate low
    xSat := TRUE;                                     // 置饱和标志 [—] / raise the saturation flag
ELSE
    FC_DL_Q15NegSat := DINT_TO_INT(diNeg);            // 界内直接转换 [Q15] / in range conversion
END_IF
END_FUNCTION

(* ---- FC_DL_Q15SqrtFloor.st ---- *)
(*
  FC_DL_Q15SqrtFloor —— Q15 定点整数平方根（逐位法），结果 Q15
  分类：DL_Base | 复杂度：2 | 轮次：R86
  开源溯源：道莅原创（clean-room 自研，纯 IEC 61131-3 通用算法），无外部代码引用
  许可证：MIT
  职责：把 Q15 输入按 Q15 语义开方（即 out = floor(sqrt(in / 32768) * 32768)）：
        先把被开方数放大 15 位成 Q30，再用逐位法（bit-by-bit）求整数平方根，结果天然是 Q15。
  契约：iIn 输入 [Q15]；返回平方根 [Q15]；负输入钳 0（置 xClamp 报告）。
  边界：① 输入钳 ≥0（负数无实数根）；② 逐位法只用整数加减与除 2 / 除 4，无浮点、无开方库依赖；
        ③ 被开方数 <= 32767 * 32768 = 1.073e9 界内；④ 零全局、零物理地址、零库件依赖。
*)
FUNCTION FC_DL_Q15SqrtFloor : INT
VAR_INPUT
    iIn : INT := 0;                   // 被开方数 [Q15] / The radicand in Q15
END_VAR
VAR_OUTPUT
    xClamp : BOOL;                    // 负输入钳零标志（信息级） [—] / The negative input clamp flag
END_VAR
VAR
    diV    : DINT;                    // 已放大 15 位的被开方数 [Q30] / The radicand scaled to Q30
    diRem  : DINT;                    // 逐位法余数 [Q30] / The remainder of the bit by bit method
    diRoot : DINT;                    // 逐位法根累加器 [Q30] / The root accumulator
    diBit  : DINT;                    // 逐位法试探位（4 的幂递减） [Q30] / The trial bit decreasing by four
END_VAR
VAR CONSTANT
    DL_QS_SC   : DINT := 32768;       // 定标因子（2^15） [-] / The Q15 scaling factor
    DL_QS_TOP  : DINT := 1073741824;  // 试探位初值 2^30 [-] / The initial trial bit
    DL_QS_Z    : DINT := 0;           // 整型零常量 [-] / The integer zero constant
    DL_QS_TWO  : DINT := 2;           // 除二常量 [-] / The divide by two constant
    DL_QS_FOUR : DINT := 4;           // 除四常量 [-] / The divide by four constant
END_VAR

xClamp := FALSE;                                      // 钳位标志预置假 / preset the clamp flag false
IF iIn < DINT_TO_INT(DL_QS_Z) THEN                    // 负输入（无实数根） / a negative input has no real root
    FC_DL_Q15SqrtFloor := DINT_TO_INT(DL_QS_Z);       // 结果钳零 [Q15] / clamp the result to zero
    xClamp := TRUE;                                   // 置钳位标志 [—] / raise the clamp flag
ELSE
    diV := INT_TO_DINT(iIn) * DL_QS_SC;               // 放大 15 位成 Q30 被开方数（界内已证） [Q30] / scale to Q30
    diRem := diV;                                     // 余数初值取被开方数 [Q30] / the initial remainder
    diRoot := DL_QS_Z;                                // 根累加器清零 [Q30] / clear the root accumulator
    diBit := DL_QS_TOP;                               // 试探位从 2^30 起 [Q30] / start from the top trial bit
    WHILE diBit > diV DO                              // 试探位降到不超被开方数（逐位法前置归一） / normalise the trial bit
        diBit := diBit / DL_QS_FOUR;                  // 试探位每次降 4 倍 [Q30] / decrease the trial bit by four
    END_WHILE
    WHILE diBit > DL_QS_Z DO                          // 主循环：16 次迭代后试探位归零 / the main loop ends at zero
        IF diRem >= (diRoot + diBit) THEN              // 余数够减 / the remainder is large enough
            diRem := diRem - diRoot - diBit;          // 扣减根与试探位 [Q30] / subtract the root and the trial bit
            diRoot := (diRoot / DL_QS_TWO) + diBit;   // 根累加器置位 [Q30] / set the root accumulator bit
        ELSE
            diRoot := diRoot / DL_QS_TWO;             // 根累加器右移一位 [Q30] / shift the root accumulator
        END_IF
        diBit := diBit / DL_QS_FOUR;                  // 试探位每次降 4 倍 [Q30] / decrease the trial bit by four
    END_WHILE
    FC_DL_Q15SqrtFloor := DINT_TO_INT(diRoot);        // 逐位法根即 Q15 结果 [Q15] / the root is the Q15 result
END_IF
END_FUNCTION

(* ---- FC_DL_Q15SubSat.st ---- *)
(*
  FC_DL_Q15SubSat —— Q15 定点减法饱和
  分类：DL_Base | 复杂度：2 | 轮次：R86
  开源溯源：道莅原创（clean-room 自研，纯 IEC 61131-3 通用算法），无外部代码引用
  许可证：MIT
  职责：Q15 域 iA - iB，中间用 DINT 承载，结果按 Q15 上下界饱和（含 -32768 边界）。
  契约：输入 iA / iB 为 Q15 操作数；返回 Q15 差；xSat 报告本拍发生饱和（信息级）。
  边界：DINT 中间量 + 上下界双判，无除法、无浮点比较；零全局、零物理地址、零库件依赖。
*)
FUNCTION FC_DL_Q15SubSat : INT
VAR_INPUT
    iA : INT := 0;                    // 被减数 A [Q15] / The minuend A in Q15
    iB : INT := 0;                    // 减数 B [Q15] / The subtrahend B in Q15
END_VAR
VAR_OUTPUT
    xSat : BOOL;                      // 饱和发生标志（信息级） [—] / The saturation flag, informational
END_VAR
VAR
    diDiff : DINT;                    // 双字中间差 [Q15] / The double word intermediate difference
END_VAR
VAR CONSTANT
    Q15_MAX : DINT := 32767;          // Q15 上界 [-] / The Q15 upper bound
    Q15_MIN : DINT := -32768;         // Q15 下界 [-] / The Q15 lower bound
END_VAR

xSat := FALSE;                                        // 饱和标志预置假 / preset the saturation flag false
diDiff := INT_TO_DINT(iA) - INT_TO_DINT(iB);          // 双字域求差（|差| <= 65535 不溢出） [Q15] / subtract in DINT
IF diDiff > Q15_MAX THEN                              // 上越界 / above the upper bound
    FC_DL_Q15SubSat := DINT_TO_INT(Q15_MAX);          // 饱和到 Q15_MAX [Q15] / saturate high
    xSat := TRUE;                                     // 置饱和标志 [—] / raise the saturation flag
ELSIF diDiff < Q15_MIN THEN                           // 下越界 / below the lower bound
    FC_DL_Q15SubSat := DINT_TO_INT(Q15_MIN);          // 饱和到 Q15_MIN [Q15] / saturate low
    xSat := TRUE;                                     // 置饱和标志 [—] / raise the saturation flag
ELSE
    FC_DL_Q15SubSat := DINT_TO_INT(diDiff);           // 界内直接转换 [Q15] / in range conversion
END_IF
END_FUNCTION

(* ---- FC_DL_RealToQ15Sat.st ---- *)
(*
  FC_DL_RealToQ15Sat —— REAL 转 Q15 定点，四舍五入加饱和，非有限值归零
  分类：DL_Base | 复杂度：1 | 轮次：R86
  开源溯源：道莅原创（clean-room 自研，纯 IEC 61131-3 通用算法），无外部代码引用
  许可证：MIT
  职责：把归一化实数 fIn（-1.0..+1.0 对应 -32768..32767）转成 Q15 整数：
        非有限值（NaN / Inf）一律归零；放大 32768 后按符号做四舍五入，再按 Q15 上下界饱和。
  契约：fIn 输入 [归一化实数 -1.0..1.0]；返回 Q15 值；xInvalid 报告输入为非有限值（信息级）。
  边界：① NaN 用自反判（fIn <> fIn）、Inf 用绝对上限判（ABS(fIn) > 1.0E30），禁用近似阈值；
        ② 实数转整前的上限兜底：放大值越 40000 时直接饱和，避免 LREAL_TO_DINT 越域未定义；
        ③ 零全局、零物理地址、零库件依赖。
*)
FUNCTION FC_DL_RealToQ15Sat : INT
VAR_INPUT
    fIn : REAL := 0.0;                // 归一化输入实数 [归一化] / The normalised real input
END_VAR
VAR_OUTPUT
    xInvalid : BOOL;                  // 输入为非有限值（信息级，已归零） [—] / The input was not finite and was zeroed
    xSat     : BOOL;                  // 越界饱和标志（信息级） [—] / The range saturation flag
END_VAR
VAR
    fScaled : LREAL;                  // 放大 32768 倍后的实数 [Q15 实数域] / The scaled real value
    diR     : DINT;                   // 四舍五入后的整数暂存 [Q15] / The rounded integer stage
END_VAR
VAR CONSTANT
    Q15_MAX    : DINT  := 32767;      // Q15 上界 [-] / The Q15 upper bound
    Q15_MIN    : DINT  := -32768;     // Q15 下界 [-] / The Q15 lower bound
    DL_QR_SC   : LREAL := 32768.0;    // 定标因子（2^15） [-] / The Q15 scaling factor
    DL_QR_HALF : LREAL := 0.5;        // 四舍五入偏置 [-] / The rounding bias
    DL_QR_LIM  : LREAL := 40000.0;    // 转整前的实数上限兜底 [-] / The real upper guard before conversion
    DL_QR_INF  : REAL  := 1.0E30;     // 非有限 / 越界判据上限 [-] / The magnitude gate for non finite detection
    DL_QR_TINY : LREAL := 1.0E-9;     // 浮点零比较容差 [-] / The floating point zero tolerance
    DL_QR_Z    : DINT  := 0;          // 整型零常量 [-] / The integer zero constant
END_VAR

xInvalid := FALSE;                                    // 非有限标志预置假 / preset the non finite flag false
xSat := FALSE;                                        // 饱和标志预置假 / preset the saturation flag false
IF (fIn <> fIn) OR (ABS(fIn) > DL_QR_INF) THEN        // 自反判 NaN 或越限判 Inf（R 规则禁用近似阈值） / NaN or Inf
    FC_DL_RealToQ15Sat := DINT_TO_INT(DL_QR_Z);       // 非有限值归零 [Q15] / zero the non finite input
    xInvalid := TRUE;                                 // 置非有限标志 [—] / raise the non finite flag
ELSE
    fScaled := REAL_TO_LREAL(fIn) * DL_QR_SC;         // 放大 32768 倍 [Q15 实数域] / scale by the Q15 factor
    IF fScaled > DL_QR_LIM THEN                       // 转整前上限兜底（正溢出） / the positive conversion guard
        FC_DL_RealToQ15Sat := DINT_TO_INT(Q15_MAX);   // 直接饱和到 Q15_MAX [Q15] / saturate high
        xSat := TRUE;                                 // 置饱和标志 [—] / raise the saturation flag
    ELSIF fScaled < -DL_QR_LIM THEN                   // 转整前下限兜底（负溢出） / the negative conversion guard
        FC_DL_RealToQ15Sat := DINT_TO_INT(Q15_MIN);   // 直接饱和到 Q15_MIN [Q15] / saturate low
        xSat := TRUE;                                 // 置饱和标志 [—] / raise the saturation flag
    ELSE
        IF fScaled >= DL_QR_HALF THEN                 // 非负做加偏置四舍五入 / non negative rounding
            diR := LREAL_TO_DINT(fScaled + DL_QR_HALF); // 加 0.5 后截断 [Q15] / add a half then truncate
        ELSIF fScaled <= -DL_QR_HALF THEN             // 非正做减偏置四舍五入 / non positive rounding
            diR := LREAL_TO_DINT(fScaled - DL_QR_HALF); // 减 0.5 后截断 [Q15] / subtract a half then truncate
        ELSE
            diR := DL_QR_Z;                           // |值| < 0.5 归零（近零带） [Q15] / the near zero band
        END_IF
        IF diR > Q15_MAX THEN                         // 上越界 / above the upper bound
            FC_DL_RealToQ15Sat := DINT_TO_INT(Q15_MAX); // 饱和到 Q15_MAX [Q15] / saturate high
            xSat := TRUE;                             // 置饱和标志 [—] / raise the saturation flag
        ELSIF diR < Q15_MIN THEN                      // 下越界 / below the lower bound
            FC_DL_RealToQ15Sat := DINT_TO_INT(Q15_MIN); // 饱和到 Q15_MIN [Q15] / saturate low
            xSat := TRUE;                             // 置饱和标志 [—] / raise the saturation flag
        ELSE
            FC_DL_RealToQ15Sat := DINT_TO_INT(diR);   // 界内直接转换 [Q15] / in range conversion
        END_IF
    END_IF
END_IF
END_FUNCTION

(* ---- FC_DL_ReverseBitsLword.st ---- *)
(*
  ==================================================================
  组件名 Component  : FC_DL_ReverseBitsLword
  分类   Category   : DL_Base
  前缀   Naming     : FC_DL_ ｜ b/n/u/f/t/e/st 类型前缀制（R265）
  复杂度 Complexity  : 低
  版本   Version    : 1.0.0
  功能   Purpose    : LWORD 64 位序整体反转（ReverseBitsWord 的 64 位域升版变体）。
  来源   Source     : t2-1-lgf-bitlogic（位逻辑族 64 位变体）
  平台   Platform   : 纯 IEC 61131-3（FOR / SHL / SHR / AND / OR），三平台通用
  分工声明 Split     : 与 FC_DL_ReverseBitsWord（32 位域属主）分工——本件只做
                      LWORD 域，不重声明低位宽件；移位量恒为 1（R48 归一纪律：
                      全程无 ≥ 位宽的移位量，无拆半区）。
  作者   Author     : 道莅代码库 · PLC 编程专家（R61）
  归属 Ownership     : 本件无 TYPE 声明；引用件类型全部 IEC 标准原生。
  ------------------------------------------------------------------
  边界 Boundary     :
                      一 uSrc = 0 → uRev = 0 且 bValid = TRUE 恒成立（全零可逆）；
                      二 反转是全域双射：任何输入都有唯一合法输出，本件无钳位、
                         无故障路径，故按 R90 反证不加任何错误码（bError 恒假、
                         eErr 恒零，属声明性常量，沿 TwoStepConfirm bError 先例）；
                      三 无状态纯函数：局部量段 1 显式预置（R254）。
  错误码   Codes    : 无（R90 反证：反转全域可逆，无任何可故障场景，不加码）。
  验收   Acceptance :
    算法已证（脚本）：未跑 ｜ 编译器已证（三平台）：未跑
    V1 uSrc=16#0000_0000_0000_0001 → uRev=16#8000_0000_0000_0000
    V2 uSrc=16#8000_0000_0000_0000 → uRev=16#0000_0000_0000_0001
    V3 uSrc=0 → uRev=0、bValid=TRUE
  修订记录 Revision  :
    2026-11-21  v1.0.0  R61 首版（批 1 · 序号 1）
  ==================================================================
*)
FUNCTION FC_DL_ReverseBitsLword : BOOL
VAR_IN_OUT
    uSrc : LWORD; // 待反转源字 [位图] / the source word to reverse
END_VAR
VAR_OUTPUT
    uRev   : LWORD;       // 反转结果字 [位图] / the reversed word
    bValid : BOOL;        // 结果可用标志（恒真：全域可逆）[-] / the validity flag, always true
    eErr   : UDINT;       // 错误码，0 = 正常（恒零：无故障路径）/ the error code, constant zero
    bError : BOOL;        // 错误标志（恒假：无故障路径，边界二）/ the error flag, constant false
END_VAR
VAR
    uWork : LWORD; // 移位工作副本（每拍右移一位耗尽）/ the shifting work copy
    k     : DINT;  // 位循环索引 [位] / the bit loop index
END_VAR

// 段 1｜返回值与输出预置（局部量显式预置，R254）/ segment 1, the preset of the return and the outputs
FC_DL_ReverseBitsLword := FALSE; // 返回值预置假 / preset the return false
uRev := 16#0000_0000_0000_0000; // 结果字预置零 / preset the result zero
bValid := FALSE; // 有效标志预置假（出口置真）/ preset the validity false
eErr := 16#0000_0000; // 错误码预置正常 / preset the code to ok
bError := FALSE; // 错误标志预置假（全域可逆，无故障路径）/ preset the error flag false
uWork := uSrc; // 工作副本装入源字 / load the work copy from the source

// 段 2｜64 位逐位反转（移位量恒 1，结构性安全于 R48）/ segment 2, the bit by bit reversal with a constant shift of one
FOR k := 0 TO 63 DO // 有界循环恰好 64 次 / the bounded loop of exactly sixty four rounds
    uRev := SHL(uRev, 1) OR (uWork AND 16#0000_0000_0000_0001); // 结果左移一位并装入源字最低位 / shift the result left and append the lowest source bit
    uWork := SHR(uWork, 1); // 源字右移一位 / shift the source right
END_FOR

// 段 3｜出口（反转全域可逆，恒成功）/ segment 3, the outlet, always successful
bValid := TRUE; // 有效标志置真 / raise the validity
FC_DL_ReverseBitsLword := TRUE; // 返回成功 / return success
END_FUNCTION

(* ---- FC_DL_RolEx.st ---- *)
(*==============================================================================
 * 组件名称 (Component)  : FC_DL_RolEx
 * 所属子库 (Sublibrary) : DL_Base
 * 当前版本 (Version)    : 1.0.0
 * 兼容性   (Platform)   : CODESYS 3.5 / TwinCAT 3 / 汇川 InoProShop / Machine Expert
 *                         仅依赖 Standard.library 的 SHL / SHR 内建函数，
 *                         循环语义由移位合成显式构造，无厂商 ROL 方言依赖
 * 功能一句话 (Summary)  : 循环左移防御包装：移位量对位宽取模归一后再循环，
 *                         杜绝平台相关行为，循环位不丢。
 * 功能描述 (Function)   : 对被移位位串按移位量 nN 循环左移。归一策略写死：
 *                         nN 先 MOD 32 归一到 0 到 31（nN 为 USINT 天然非负，
 *                         禁用 MOD 对负数的平台歧义取余的前提由类型系统保证）；
 *                         归一后 nN = 0 直接返回原值（整圈等价于不动，不置码）；
 *                         归一后 1 到 31 用「左移 nN OR 右移 (32 − nN)」位合成
 *                         构造循环语义，两个合成移位量均严格落在 1 到 31 安全域。
 * 溯源     (Origin)     : IEC 61131-3 标准语义的道莅防御性实现
 *                         （接口语义由 IEC 61131-3 定义，clean-room 重写，
 *                         参考公开标准条款）
 * 支持位宽 (Width Note) : 本件按 DWORD（32 位）主类型实现，仅支持 32 位位串；
 *                         BYTE / WORD 调用方先显式转换到 DWORD 后调用，再按需
 *                         截回原位宽（头注释显式声明，不做 ANY_BIT 泛型）。
 * 类型裁定 (Type Note)  : 码位段 16#0001_xxxx 为全库共享 32 位段，WORD 容量不足，
 *                         故 uDiag 采用 UDINT 承载（与库内 uErrorId : UDINT 惯例一致）
 * 依赖     (Depends)    : 无 DL_ 内部依赖；Standard.library: SHL / SHR
 * 红线自检 (Redline)    : R1 ✓ 零全局变量与外部变量引用 ｜ R2 ✓ 零物理 IO 地址直写
 *                         R3 ✓ 纯 IEC 61131-3 ｜ R4 ✓ 移位量 MOD 归一（合成移位
 *                         量恒在 1 到 31 安全域）｜ R5 ✓ 全变量中英双语同行注释
 *                         R6 N/A（纯函数，无 CASE/ENUM 状态机，按批 1 口径标 N/A）
 *                         R7 N/A（FC 为纯函数，无实例调用，头注释显式说明）
 * 防御行为声明 (Defense): ① 归一先行：nN ≥ 32 时先 MOD 32 归一并置信息码
 *                           16#0001_0158（已归一提示），归一后绝不出现 ≥ 位宽
 *                           的移位量，杜绝平台对超宽循环移位的歧义行为；
 *                         ② nN 为 USINT 类型天然非负，MOD 只作用于非负域，
 *                           负数取余的平台歧义（如商向零取整方向不一）从类型
 *                           系统层面被排除，该前提已在头注释写死；
 *                         ③ 归一后 nN = 0 直接返回原值且不置码（整圈无事件）；
 *                         ④ 位合成用「SHL(uIn, nN) OR SHR(uIn, 32 − nN)」，
 *                           nN 归一后为 1 到 31，故 32 − nN 恒为 1 到 31，
 *                           两个移位量均不触碰「移位量 = 位宽」禁区，循环位不丢；
 *                         ⑤ 32（位宽）提为只读常量，禁魔法数。
 * 修订历史 (Revision)   :
 *   2026-11-16  v1.0.0  首版入库（R14 批 3 · T0 快车道）
 *============================================================================*)
FUNCTION FC_DL_RolEx : DWORD
VAR_INPUT
    uIn : DWORD;   // 被循环移位位串 [位] / Bit string to be rotated
    nN  : USINT;   // 移位量 [bit]，USINT 天然非负，MOD 仅作用于非负域 / Shift amount [bit], USINT is non-negative, MOD applied on the non-negative domain only
END_VAR
VAR_OUTPUT
    uDiag : UDINT; // 诊断字，16#0001_0158=移位量已 MOD 32 归一，0=无事件 / Diag word, 16#0001_0158=shift amount reduced by MOD 32, 0=no event
END_VAR
VAR
    nNorm : USINT; // 归一后移位量 [bit]，域 0 到 31 / Normalized shift amount [bit], range 0 to 31
END_VAR
VAR CONSTANT
    DL_RO_WIDTH : USINT := 32;  // 位宽常量 [bit]，MOD 归一与合成移位共用 / Width constant [bit], shared by MOD normalization and composite shifts
END_VAR

(*------------------------------------------------------------------------------
 * 段 1｜输出与诊断预置：先归零，任何路径都不会留下脏诊断
 *      Pre-set the output and diag so no path ever leaves a stale diag
 *-----------------------------------------------------------------------------*)
FC_DL_RolEx := 16#0000_0000;   // 返回值预置全零 [位串] / Preset return value to all zero
uDiag       := 16#0000_0000;   // 诊断字预置无事件 / Preset diag word to no event
nNorm       := 0;              // 归一移位量预置 [bit] / Preset normalized shift to zero [bit]

(*------------------------------------------------------------------------------
 * 段 2｜移位量归一（防御声明①②）：nN MOD 32 归一到 0 到 31；
 *      nN 为 USINT 非负域，MOD 结果即数学取模，无负数取余歧义；
 *      nN ≥ 32 置信息码提示已归一（归一是正常防御行为，非故障）
 *      Shift-amount normalization (defense notes 1 and 2): nN MOD 32 reduces
 *      to 0 to 31; a reduction raises the informational code, not a fault
 *-----------------------------------------------------------------------------*)
IF nN >= DL_RO_WIDTH THEN
    nNorm := nN MOD DL_RO_WIDTH;   // 超宽归一：MOD 32 取模 [bit] / Oversized normalization: MOD 32 [bit]
    uDiag := 16#0001_0158;         // 信息码：移位量已 MOD 32 归一 / Informational: shift amount reduced by MOD 32
ELSE
    nNorm := nN;                   // 域内直通 [bit] / In-domain pass-through [bit]
END_IF

(*------------------------------------------------------------------------------
 * 段 3｜循环移位主体（防御声明③④）：归一后 0 整圈直通原值；
 *      1 到 31 用左移与右移位合成，合成移位量恒在安全域，循环位不丢
 *      Rotation body (defense notes 3 and 4): normalized zero returns as is;
 *      one to thirty one composes SHL and SHR, both amounts stay in the safe
 *      domain so no bit is ever lost
 *-----------------------------------------------------------------------------*)
IF nNorm = 0 THEN
    FC_DL_RolEx := uIn;   // 整圈（或 0 位）等价于原值直通 [位串] / A full turn (or zero shift) returns the input unchanged
ELSE
    FC_DL_RolEx := SHL(uIn, nNorm) OR SHR(uIn, DL_RO_WIDTH - nNorm);   // 位合成循环左移 [位串] / Composite rotate left
END_IF
END_FUNCTION

(* ---- FC_DL_RolLwordEx.st ---- *)
(*
    FC_DL_RolLwordEx —— LWORD 循环左移（MOD 64 归一）
    ------------------------------------------------------------------
    分类      : DL_Base / BitString
    前缀      : FC_DL_
    版本      : 1.0.0
    溯源      : IEC 61131-3 标准语义的道莅防御性实现
                （接口语义由 IEC 61131-3 定义，内部委托平台内建 ROL，
                  外围统一错误码 / 钳位 / 双语文档；clean-room 重写，
                  未复制任何闭源厂商源码，参考实现仅限 MIT/Apache 许可）
    平台      : 纯 IEC 61131-3，CODESYS / TwinCAT / InoProShop 通用
    作者      : 道莅代码库 · PLC编程专家（R17）
    ------------------------------------------------------------------
    功能说明  : LWORD 位串循环左移防御包装：移位量 nN 大于等于 64（位宽）时按 MOD 64 归一，
                并置信息级 16#0001_020A（循环移位对位宽取模仍等价，故归一而非置零——
                与左移/右移件的「超宽置零」口径刻意相反，二者语义不可混用）；
                归一后移位量为 0 时直接输出原值，不调用内建 ROL（规避零移位量的平台差异）；
                域内委托平台内建 ROL，不重实现移位内核；
                MOD 除子为常量 64（编译期恒非零），结构性满足除法前判除子非零红线；
                钳位方向：移位量按位宽取模归一（0~63），结果位宽严格保持 64 位。
    错误码    : 16#0001_020A 移位量 ≥ 64（位宽），已按 MOD 64 归一——信息级，正常防御
                16#0001_020B 预留禁用（信息级，不得挪用）
                16#0001_02FD 预留禁用（故障级，不得挪用）
                16#0001_02FE 预留禁用（故障级，不得挪用）
                16#0001_02FF 预留禁用（故障级，不得挪用）
    状态机    : R6 标注 N/A —— 本组件为纯函数无顺序状态机，无 CASE 可写，非法状态不可能出现，故以本节说明替代 ELSE 兜底
    修订记录  : 2026-11-16 v1.0.0 首次入库（R17）
*)
FUNCTION FC_DL_RolLwordEx : LWORD
VAR_INPUT
    uIn : LWORD; // 被循环移位位串 [位] / bit string to be rotated [bit]
    nN  : USINT; // 循环移位量 [bit]，USINT 天然非负，范围 0~255 / rotate amount [bit], USINT is non-negative by type, range 0..255
END_VAR
VAR_OUTPUT
    eErr   : UDINT; // 错误码，0=正常 / error id, 0=ok
    bError : BOOL;  // 是否出错，eErr 非 0 时为 TRUE / error flag, TRUE when eErr is nonzero
    bValid : BOOL;  // 输出是否有效可用 / output valid flag
END_VAR
VAR CONSTANT
    DL_LW_WIDTH : USINT := 64; // LWORD 位宽常量，兼作 MOD 除子（编译期恒非零） [bit] / LWORD width constant, also the MOD divisor, never zero [bit]
END_VAR
VAR
    nShift : USINT; // 归一后的实际移位量 0~63 [bit] / normalized shift amount 0..63 [bit]
END_VAR

// 段 1｜输出与错误状态预置 / segment 1, preset output and error status
FC_DL_RolLwordEx := uIn; // 输出预置为原值（零移位等价语义），任何路径不留脏值 [位串] / preset output to the input, the zero-shift identity, no stale value on any path [bit string]
eErr   := 0;     // 预置无错误 / preset no error
bError := FALSE; // 预置无故障（本件无故障级路径） / preset no fault, no fault-level path here
bValid := FALSE; // 预置输出无效，通过归一后置位 / preset invalid, set TRUE after normalization

// 段 2｜移位量归一（MOD 位宽） / segment 2, shift amount normalization (modulo width)
nShift := nN; // 默认按原移位量直通 [bit] / pass the original shift amount through by default [bit]
IF nN >= DL_LW_WIDTH THEN // 循环移位对位宽取模仍等价，故归一而非置零 [bit] / rotate modulo the width stays equivalent, so normalize instead of zeroing [bit]
    nShift := nN MOD DL_LW_WIDTH; // 除子为编译期常量 64，恒非零 [bit] / divisor is the compile-time constant 64, never zero [bit]
    eErr := 16#0001_020A;         // 信息级：移位量已归一，正常防御 / info level: shift amount normalized, normal defence
ELSE
    eErr := 0;                    // 未超宽，无记录 / not oversized, nothing recorded
END_IF

// 段 3｜零移位量与域内委托循环移位（末段） / segment 3, zero-shift pass-through and in-domain delegated rotate (final)
IF nShift = 0 THEN
    FC_DL_RolLwordEx := uIn; // 零移位量直接输出原值，规避内建 ROL 的平台差异 [位串] / zero shift passes the input through, avoiding platform differences of built-in ROL [bit string]
ELSE
    FC_DL_RolLwordEx := ROL(uIn, nShift); // 域内委托平台内建 ROL，不重实现移位内核 [位串] / in-domain delegate to built-in ROL, shift kernel not re-implemented [bit string]
END_IF
bError := FALSE; // 信息级不置故障 / info level never raises fault
bValid := TRUE;  // 归一后输出有效可用 / output is valid after normalization
END_FUNCTION
